(* IEC 61131-3 sources: plc-st-coding-agent/progress/evidence/f14_v14_remaining_20261113/jobs/codex_deepseek-v4pro (part 2) *)

(* ---- public-hard-01.raw_candidate_03.st ---- *)
(* CONTRACT_RULES [] *)

(* ENGINEERING_CONTRACT
   - ESTOP: ESTOP=FALSE forces every output OFF in this scan; manual and auto commands are inhibited.
   - Manual runs: only while OpeMode=FALSE and ESTOP=TRUE; each start button rising edge toggles its retained output latch.
   - Auto sequence: AUTOSTART rising edge while OpeMode=TRUE enters FILL_A; output valves follow the sequence below.
   - Valve A: ON in FILL_A; Level>=50 closes A and opens B (PUB012).
   - Valve B: ON in FILL_B; Level>=80 closes B (PUB012/PUB013).
   - ProcessMode=FALSE: at Level>=80 mixer starts; MixMotorComplete latches completion, then mixer off and Valve D ON, sequence done (PUB014).
   - ProcessMode=TRUE: at Level>=80 Valve C opens; Level>=100 closes C and starts mixer; completion opens D (PUB014).
   - Mix complete is latched until the next AUTOSTART; Valve D remains ON in DONE because no stop/reset is stated.
   - Thresholds are inclusive >=; Level is INT cm; PROCESSMODE is read live at the 80 cm transition.
*)

TYPE E_MaterialProportioningState :
(
    MP_IDLE,
    MP_FILL_A,
    MP_FILL_B,
    MP_MIX_SIMPLE,
    MP_FILL_C,
    MP_MIX_C,
    MP_DONE
) := MP_IDLE;
END_TYPE;

FUNCTION_BLOCK MaterialProportioningControl
VAR_INPUT
    estop : BOOL;
    opeMode : BOOL;
    valveAStart : BOOL;
    valveBStart : BOOL;
    valveCStart : BOOL;
    valveDStart : BOOL;
    mixMotorStart : BOOL;
    autoStart : BOOL;
    processMode : BOOL;
    levelSensor : INT;
    mixMotorComplete : BOOL;
END_VAR
VAR_OUTPUT
    valveARun : BOOL;
    valveBRun : BOOL;
    valveCRun : BOOL;
    valveDRun : BOOL;
    mixMotorRun : BOOL;
END_VAR
VAR
    tmp_trigValveA : R_TRIG;
    tmp_trigValveB : R_TRIG;
    tmp_trigValveC : R_TRIG;
    tmp_trigValveD : R_TRIG;
    tmp_trigMixMotor : R_TRIG;
    tmp_trigAutoStart : R_TRIG;

    manualValveARun : BOOL := FALSE;
    manualValveBRun : BOOL := FALSE;
    manualValveCRun : BOOL := FALSE;
    manualValveDRun : BOOL := FALSE;
    manualMixMotorRun : BOOL := FALSE;

    state : E_MaterialProportioningState := MP_IDLE;
    mixCompleteLatched : BOOL := FALSE;
END_VAR

tmp_trigValveA(CLK := valveAStart);
tmp_trigValveB(CLK := valveBStart);
tmp_trigValveC(CLK := valveCStart);
tmp_trigValveD(CLK := valveDStart);
tmp_trigMixMotor(CLK := mixMotorStart);
tmp_trigAutoStart(CLK := autoStart);

IF NOT estop THEN
    valveARun := FALSE;
    valveBRun := FALSE;
    valveCRun := FALSE;
    valveDRun := FALSE;
    mixMotorRun := FALSE;

ELSIF NOT opeMode THEN
    state := MP_IDLE;
    mixCompleteLatched := FALSE;

    IF tmp_trigValveA.Q THEN
        manualValveARun := NOT manualValveARun;
    END_IF;
    IF tmp_trigValveB.Q THEN
        manualValveBRun := NOT manualValveBRun;
    END_IF;
    IF tmp_trigValveC.Q THEN
        manualValveCRun := NOT manualValveCRun;
    END_IF;
    IF tmp_trigValveD.Q THEN
        manualValveDRun := NOT manualValveDRun;
    END_IF;
    IF tmp_trigMixMotor.Q THEN
        manualMixMotorRun := NOT manualMixMotorRun;
    END_IF;

    valveARun := manualValveARun;
    valveBRun := manualValveBRun;
    valveCRun := manualValveCRun;
    valveDRun := manualValveDRun;
    mixMotorRun := manualMixMotorRun;

ELSE
    IF tmp_trigAutoStart.Q THEN
        state := MP_FILL_A;
        mixCompleteLatched := FALSE;
    END_IF;

    CASE state OF
        MP_IDLE:
            valveARun := FALSE;
            valveBRun := FALSE;
            valveCRun := FALSE;
            valveDRun := FALSE;
            mixMotorRun := FALSE;

        MP_FILL_A:
            valveARun := TRUE;
            valveBRun := FALSE;
            valveCRun := FALSE;
            valveDRun := FALSE;
            mixMotorRun := FALSE;

            IF levelSensor >= 80 THEN
                valveARun := FALSE;
                valveBRun := FALSE;
                IF NOT processMode THEN
                    mixMotorRun := TRUE;
                    mixCompleteLatched := FALSE;
                    state := MP_MIX_SIMPLE;
                ELSIF levelSensor >= 100 THEN
                    valveCRun := FALSE;
                    mixMotorRun := TRUE;
                    mixCompleteLatched := FALSE;
                    state := MP_MIX_C;
                ELSE
                    valveCRun := TRUE;
                    state := MP_FILL_C;
                END_IF;
            ELSIF levelSensor >= 50 THEN
                valveARun := FALSE;
                valveBRun := TRUE;
                state := MP_FILL_B;
            END_IF;

        MP_FILL_B:
            valveARun := FALSE;
            valveBRun := TRUE;
            valveCRun := FALSE;
            valveDRun := FALSE;
            mixMotorRun := FALSE;

            IF levelSensor >= 80 THEN
                valveBRun := FALSE;
                IF NOT processMode THEN
                    mixMotorRun := TRUE;
                    mixCompleteLatched := FALSE;
                    state := MP_MIX_SIMPLE;
                ELSE
                    IF levelSensor >= 100 THEN
                        valveCRun := FALSE;
                        mixMotorRun := TRUE;
                        mixCompleteLatched := FALSE;
                        state := MP_MIX_C;
                    ELSE
                        valveCRun := TRUE;
                        state := MP_FILL_C;
                    END_IF;
                END_IF;
            END_IF;

        MP_FILL_C:
            valveARun := FALSE;
            valveBRun := FALSE;
            valveCRun := TRUE;
            valveDRun := FALSE;
            mixMotorRun := FALSE;

            IF levelSensor >= 100 THEN
                valveCRun := FALSE;
                mixMotorRun := TRUE;
                mixCompleteLatched := FALSE;
                state := MP_MIX_C;
            END_IF;

        MP_MIX_SIMPLE:
            valveARun := FALSE;
            valveBRun := FALSE;
            valveCRun := FALSE;
            valveDRun := FALSE;
            mixMotorRun := TRUE;

            IF mixMotorComplete THEN
                mixCompleteLatched := TRUE;
            END_IF;

            IF mixCompleteLatched THEN
                mixMotorRun := FALSE;
                valveDRun := TRUE;
                state := MP_DONE;
            END_IF;

        MP_MIX_C:
            valveARun := FALSE;
            valveBRun := FALSE;
            valveCRun := FALSE;
            valveDRun := FALSE;
            mixMotorRun := TRUE;

            IF mixMotorComplete THEN
                mixCompleteLatched := TRUE;
            END_IF;

            IF mixCompleteLatched THEN
                mixMotorRun := FALSE;
                valveDRun := TRUE;
                state := MP_DONE;
            END_IF;

        MP_DONE:
            valveARun := FALSE;
            valveBRun := FALSE;
            valveCRun := FALSE;
            valveDRun := TRUE;
            mixMotorRun := FALSE;
    END_CASE;
END_IF;
END_FUNCTION_BLOCK

(* ---- public-hard-02.candidate_01.st ---- *)
(*
ENGINEERING_CONTRACT
- conveyorLeft | activation: ST_MOVING and target<current | hold: while ST_MOVING | reset: target sensor arrival or non-moving state | same-scan: final settled state/target controls write | PUB001,PUB005.
- conveyorRight | activation: ST_MOVING and target>current | hold: while ST_MOVING | reset: target sensor arrival or non-moving state | same-scan: final settled state/target controls write | PUB001,PUB005.
- local_state | activation: ST_IDLE+start -> ST_MOVING; ST_MOVING+sensor -> ST_WAIT_COMPLETION/ST_DONE/next ST_MOVING; ST_WAIT_COMPLETION+completion -> ST_MOVING/ST_DONE | hold: retained every scan | reset/deactivation: above transitions | same-scan: inputs iterated to fixed point before outputs | units: seq index 1..processLength, stations 1..5 | PUB001-PUB005.
- local_step_index/current/target | update: start, sensor, completion | hold: otherwise | bounds: step 1..8, current/target 1..5 | PUB002,PUB005.
- Direction rule: one target per step yields exactly one direction output; equal/unknown target de-energizes both.
- Unspecified: no restart/reset after station5; completion signals treated as levels.
*)
(* CONTRACT_RULES [] *)

TYPE CONTROL_STATE :
(
    ST_IDLE,
    ST_MOVING,
    ST_WAIT_COMPLETION,
    ST_DONE
);
END_TYPE;

FUNCTION_BLOCK FlexibleProcessingControl
VAR_INPUT
    processLength : USINT;
    sensor1 : BOOL;
    sensor2 : BOOL;
    sensor3 : BOOL;
    sensor4 : BOOL;
    sensor5 : BOOL;
    station1Start : BOOL;
    station2Complete : BOOL;
    station3Complete : BOOL;
    station4Complete : BOOL;
    processSequence : ARRAY[1..8] OF USINT;
END_VAR
VAR_OUTPUT
    conveyorLeft : BOOL;
    conveyorRight : BOOL;
END_VAR
VAR
    local_state : CONTROL_STATE := ST_IDLE;
    local_step_index : USINT := 0;
    local_current_station : USINT := 1;
    local_target_station : USINT := 0;
    local_completion_active : BOOL := FALSE;
    local_target_sensor_active : BOOL := FALSE;
    local_fixpoint_scan : INT := 0;
    local_fixpoint_stable : BOOL := FALSE;
END_VAR

FOR local_fixpoint_scan := 1 TO 20 DO
    local_fixpoint_stable := TRUE;

    local_completion_active := FALSE;
    IF local_target_station = 2 THEN
        local_completion_active := station2Complete;
    ELSIF local_target_station = 3 THEN
        local_completion_active := station3Complete;
    ELSIF local_target_station = 4 THEN
        local_completion_active := station4Complete;
    END_IF;

    local_target_sensor_active := FALSE;
    IF local_target_station = 2 THEN
        local_target_sensor_active := sensor2;
    ELSIF local_target_station = 3 THEN
        local_target_sensor_active := sensor3;
    ELSIF local_target_station = 4 THEN
        local_target_sensor_active := sensor4;
    ELSIF local_target_station = 5 THEN
        local_target_sensor_active := sensor5;
    END_IF;

    CASE local_state OF
        ST_IDLE:
            IF sensor1 AND station1Start THEN
                local_step_index := 1;
                local_current_station := 1;
                local_target_station := processSequence[1];
                local_state := ST_MOVING;
                local_fixpoint_stable := FALSE;
            END_IF;

        ST_MOVING:
            IF local_target_sensor_active THEN
                local_current_station := local_target_station;

                IF local_target_station = 5 THEN
                    local_state := ST_DONE;
                ELSIF local_completion_active THEN
                    IF local_step_index < processLength THEN
                        local_step_index := local_step_index + 1;
                        local_target_station := processSequence[local_step_index];
                        local_state := ST_MOVING;
                    ELSE
                        local_state := ST_DONE;
                    END_IF;
                ELSE
                    local_state := ST_WAIT_COMPLETION;
                END_IF;

                local_fixpoint_stable := FALSE;
            END_IF;

        ST_WAIT_COMPLETION:
            IF local_completion_active THEN
                IF local_step_index < processLength THEN
                    local_step_index := local_step_index + 1;
                    local_target_station := processSequence[local_step_index];
                    local_state := ST_MOVING;
                ELSE
                    local_state := ST_DONE;
                END_IF;

                local_fixpoint_stable := FALSE;
            END_IF;

        ST_DONE:
            local_fixpoint_stable := TRUE;
    END_CASE;

    IF local_fixpoint_stable THEN
        EXIT;
    END_IF;
END_FOR;

IF local_state = ST_MOVING THEN
    IF local_target_station > local_current_station THEN
        conveyorLeft := FALSE;
        conveyorRight := TRUE;
    ELSIF local_target_station < local_current_station THEN
        conveyorLeft := TRUE;
        conveyorRight := FALSE;
    ELSE
        conveyorLeft := FALSE;
        conveyorRight := FALSE;
    END_IF;
ELSE
    conveyorLeft := FALSE;
    conveyorRight := FALSE;
END_IF;

END_FUNCTION_BLOCK

(* ---- public-hard-02.candidate_02.st ---- *)
(*
ENGINEERING_CONTRACT
- conveyorLeft | activation: ST_MOVING and target<current | hold: while ST_MOVING | reset: target sensor arrival or non-moving state | same-scan: final settled state/target controls write | PUB001,PUB005.
- conveyorRight | activation: ST_MOVING and target>current | hold: while ST_MOVING | reset: target sensor arrival or non-moving state | same-scan: final settled state/target controls write | PUB001,PUB005.
- local_state | activation: ST_IDLE+start -> ST_MOVING; ST_MOVING+sensor -> ST_WAIT_COMPLETION/ST_DONE/next ST_MOVING; ST_WAIT_COMPLETION+completion -> ST_MOVING/ST_DONE | hold: retained every scan | reset/deactivation: above transitions | same-scan: inputs iterated to fixed point before outputs | units: seq index 1..processLength, stations 1..5 | PUB001-PUB005.
- local_step_index/current/target | update: start, sensor, completion | hold: otherwise | bounds: step 1..8, current/target 1..5 | PUB002,PUB005.
- Direction rule: one target per step yields exactly one direction output; equal/unknown target de-energizes both.
- Unspecified: completion signals treated as levels; ST_DONE restarts on sensor1 AND station1Start.
*)
(* CONTRACT_RULES [] *)

TYPE CONTROL_STATE :
(
    ST_IDLE,
    ST_MOVING,
    ST_WAIT_COMPLETION,
    ST_DONE
);
END_TYPE;

FUNCTION_BLOCK FlexibleProcessingControl
VAR_INPUT
    processLength : USINT;
    sensor1 : BOOL;
    sensor2 : BOOL;
    sensor3 : BOOL;
    sensor4 : BOOL;
    sensor5 : BOOL;
    station1Start : BOOL;
    station2Complete : BOOL;
    station3Complete : BOOL;
    station4Complete : BOOL;
    processSequence : ARRAY[1..8] OF USINT;
END_VAR
VAR_OUTPUT
    conveyorLeft : BOOL;
    conveyorRight : BOOL;
END_VAR
VAR
    local_state : CONTROL_STATE := ST_IDLE;
    local_step_index : USINT := 0;
    local_current_station : USINT := 1;
    local_target_station : USINT := 0;
    local_completion_active : BOOL := FALSE;
    local_target_sensor_active : BOOL := FALSE;
    local_fixpoint_scan : INT := 0;
    local_fixpoint_stable : BOOL := FALSE;
END_VAR

FOR local_fixpoint_scan := 1 TO 20 DO
    local_fixpoint_stable := TRUE;

    local_completion_active := FALSE;
    IF local_target_station = 2 THEN
        local_completion_active := station2Complete;
    ELSIF local_target_station = 3 THEN
        local_completion_active := station3Complete;
    ELSIF local_target_station = 4 THEN
        local_completion_active := station4Complete;
    END_IF;

    local_target_sensor_active := FALSE;
    IF local_target_station = 2 THEN
        local_target_sensor_active := sensor2;
    ELSIF local_target_station = 3 THEN
        local_target_sensor_active := sensor3;
    ELSIF local_target_station = 4 THEN
        local_target_sensor_active := sensor4;
    ELSIF local_target_station = 5 THEN
        local_target_sensor_active := sensor5;
    END_IF;

    CASE local_state OF
        ST_IDLE:
            IF sensor1 AND station1Start THEN
                local_step_index := 1;
                local_current_station := 1;
                local_target_station := processSequence[1];
                local_state := ST_MOVING;
                local_fixpoint_stable := FALSE;
            END_IF;

        ST_MOVING:
            IF local_target_sensor_active THEN
                local_current_station := local_target_station;

                IF local_target_station = 5 THEN
                    local_state := ST_DONE;
                ELSIF local_completion_active THEN
                    IF local_step_index < processLength THEN
                        local_step_index := local_step_index + 1;
                        local_target_station := processSequence[local_step_index];
                        local_state := ST_MOVING;
                    ELSE
                        local_state := ST_DONE;
                    END_IF;
                ELSE
                    local_state := ST_WAIT_COMPLETION;
                END_IF;

                local_fixpoint_stable := FALSE;
            END_IF;

        ST_WAIT_COMPLETION:
            IF local_completion_active THEN
                IF local_step_index < processLength THEN
                    local_step_index := local_step_index + 1;
                    local_target_station := processSequence[local_step_index];
                    local_state := ST_MOVING;
                ELSE
                    local_state := ST_DONE;
                END_IF;

                local_fixpoint_stable := FALSE;
            END_IF;

        ST_DONE:
            IF sensor1 AND station1Start THEN
                local_step_index := 1;
                local_current_station := 1;
                local_target_station := processSequence[1];
                local_state := ST_MOVING;
                local_fixpoint_stable := FALSE;
            END_IF;
    END_CASE;

    IF local_fixpoint_stable THEN
        EXIT;
    END_IF;
END_FOR;

IF local_state = ST_MOVING THEN
    IF local_target_station > local_current_station THEN
        conveyorLeft := FALSE;
        conveyorRight := TRUE;
    ELSIF local_target_station < local_current_station THEN
        conveyorLeft := TRUE;
        conveyorRight := FALSE;
    ELSE
        conveyorLeft := FALSE;
        conveyorRight := FALSE;
    END_IF;
ELSE
    conveyorLeft := FALSE;
    conveyorRight := FALSE;
END_IF;

END_FUNCTION_BLOCK

(* ---- public-hard-02.candidate_03.st ---- *)
(*
ENGINEERING_CONTRACT
- conveyorLeft | activation: ST_MOVING and target<current | hold: while ST_MOVING | reset: target sensor arrival or non-moving state | same-scan: final settled state/target controls write | PUB001,PUB005.
- conveyorRight | activation: ST_MOVING and target>current | hold: while ST_MOVING | reset: target sensor arrival or non-moving state | same-scan: final settled state/target controls write | PUB001,PUB005.
- local_state | activation: ST_IDLE+start -> ST_MOVING; ST_MOVING+sensor -> ST_WAIT_COMPLETION/ST_DONE/next ST_MOVING; ST_WAIT_COMPLETION+completion -> ST_MOVING/ST_DONE | hold: retained every scan | reset/deactivation: above transitions | same-scan: one transition per scan based on current public inputs | units: seq index 1..processLength, stations 1..5 | PUB001-PUB005.
- local_step_index/current/target | update: start, sensor, completion | hold: otherwise | bounds: step 1..8, current/target 1..5 | PUB002,PUB005.
- Direction rule: one target per step yields exactly one direction output; equal/unknown target de-energizes both.
- Unspecified: completion signals treated as levels; ST_DONE restarts on sensor1 AND station1Start.
*)
(* CONTRACT_RULES [] *)

TYPE CONTROL_STATE :
(
    ST_IDLE,
    ST_MOVING,
    ST_WAIT_COMPLETION,
    ST_DONE
);
END_TYPE;

FUNCTION_BLOCK FlexibleProcessingControl
VAR_INPUT
    processLength : USINT;
    sensor1 : BOOL;
    sensor2 : BOOL;
    sensor3 : BOOL;
    sensor4 : BOOL;
    sensor5 : BOOL;
    station1Start : BOOL;
    station2Complete : BOOL;
    station3Complete : BOOL;
    station4Complete : BOOL;
    processSequence : ARRAY[1..8] OF USINT;
END_VAR
VAR_OUTPUT
    conveyorLeft : BOOL;
    conveyorRight : BOOL;
END_VAR
VAR
    local_state : CONTROL_STATE := ST_IDLE;
    local_step_index : USINT := 0;
    local_current_station : USINT := 1;
    local_target_station : USINT := 0;
    local_completion_active : BOOL := FALSE;
    local_target_sensor_active : BOOL := FALSE;
END_VAR

    local_completion_active := FALSE;
    IF local_target_station = 2 THEN
        local_completion_active := station2Complete;
    ELSIF local_target_station = 3 THEN
        local_completion_active := station3Complete;
    ELSIF local_target_station = 4 THEN
        local_completion_active := station4Complete;
    END_IF;

    local_target_sensor_active := FALSE;
    IF local_target_station = 2 THEN
        local_target_sensor_active := sensor2;
    ELSIF local_target_station = 3 THEN
        local_target_sensor_active := sensor3;
    ELSIF local_target_station = 4 THEN
        local_target_sensor_active := sensor4;
    ELSIF local_target_station = 5 THEN
        local_target_sensor_active := sensor5;
    END_IF;

    CASE local_state OF
        ST_IDLE:
            IF sensor1 AND station1Start THEN
                local_step_index := 1;
                local_current_station := 1;
                local_target_station := processSequence[1];
                local_state := ST_MOVING;
            END_IF;

        ST_MOVING:
            IF local_target_sensor_active THEN
                local_current_station := local_target_station;

                IF local_target_station = 5 THEN
                    local_state := ST_DONE;
                ELSIF local_completion_active THEN
                    IF local_step_index < processLength THEN
                        local_step_index := local_step_index + 1;
                        local_target_station := processSequence[local_step_index];
                        local_state := ST_MOVING;
                    ELSE
                        local_state := ST_DONE;
                    END_IF;
                ELSE
                    local_state := ST_WAIT_COMPLETION;
                END_IF;
            END_IF;

        ST_WAIT_COMPLETION:
            IF local_completion_active THEN
                IF local_step_index < processLength THEN
                    local_step_index := local_step_index + 1;
                    local_target_station := processSequence[local_step_index];
                    local_state := ST_MOVING;
                ELSE
                    local_state := ST_DONE;
                END_IF;
            END_IF;

        ST_DONE:
            IF sensor1 AND station1Start THEN
                local_step_index := 1;
                local_current_station := 1;
                local_target_station := processSequence[1];
                local_state := ST_MOVING;
            END_IF;
    END_CASE;

IF local_state = ST_MOVING THEN
    IF local_target_station > local_current_station THEN
        conveyorLeft := FALSE;
        conveyorRight := TRUE;
    ELSIF local_target_station < local_current_station THEN
        conveyorLeft := TRUE;
        conveyorRight := FALSE;
    ELSE
        conveyorLeft := FALSE;
        conveyorRight := FALSE;
    END_IF;
ELSE
    conveyorLeft := FALSE;
    conveyorRight := FALSE;
END_IF;

END_FUNCTION_BLOCK

(* ---- public-hard-02.patch_base_02.st ---- *)
(*
ENGINEERING_CONTRACT
- conveyorLeft | activation: ST_MOVING and target<current | hold: while ST_MOVING | reset: target sensor arrival or non-moving state | same-scan: final settled state/target controls write | PUB001,PUB005.
- conveyorRight | activation: ST_MOVING and target>current | hold: while ST_MOVING | reset: target sensor arrival or non-moving state | same-scan: final settled state/target controls write | PUB001,PUB005.
- local_state | activation: ST_IDLE+start -> ST_MOVING; ST_MOVING+sensor -> ST_WAIT_COMPLETION/ST_DONE/next ST_MOVING; ST_WAIT_COMPLETION+completion -> ST_MOVING/ST_DONE | hold: retained every scan | reset/deactivation: above transitions | same-scan: inputs iterated to fixed point before outputs | units: seq index 1..processLength, stations 1..5 | PUB001-PUB005.
- local_step_index/current/target | update: start, sensor, completion | hold: otherwise | bounds: step 1..8, current/target 1..5 | PUB002,PUB005.
- Direction rule: one target per step yields exactly one direction output; equal/unknown target de-energizes both.
- Unspecified: no restart/reset after station5; completion signals treated as levels.
*)
(* CONTRACT_RULES [] *)

TYPE CONTROL_STATE :
(
    ST_IDLE,
    ST_MOVING,
    ST_WAIT_COMPLETION,
    ST_DONE
);
END_TYPE;

FUNCTION_BLOCK FlexibleProcessingControl
VAR_INPUT
    processLength : USINT;
    sensor1 : BOOL;
    sensor2 : BOOL;
    sensor3 : BOOL;
    sensor4 : BOOL;
    sensor5 : BOOL;
    station1Start : BOOL;
    station2Complete : BOOL;
    station3Complete : BOOL;
    station4Complete : BOOL;
    processSequence : ARRAY[1..8] OF USINT;
END_VAR
VAR_OUTPUT
    conveyorLeft : BOOL;
    conveyorRight : BOOL;
END_VAR
VAR
    local_state : CONTROL_STATE := ST_IDLE;
    local_step_index : USINT := 0;
    local_current_station : USINT := 1;
    local_target_station : USINT := 0;
    local_completion_active : BOOL := FALSE;
    local_target_sensor_active : BOOL := FALSE;
    local_fixpoint_scan : INT := 0;
    local_fixpoint_stable : BOOL := FALSE;
END_VAR

FOR local_fixpoint_scan := 1 TO 20 DO
    local_fixpoint_stable := TRUE;

    local_completion_active := FALSE;
    IF local_target_station = 2 THEN
        local_completion_active := station2Complete;
    ELSIF local_target_station = 3 THEN
        local_completion_active := station3Complete;
    ELSIF local_target_station = 4 THEN
        local_completion_active := station4Complete;
    END_IF;

    local_target_sensor_active := FALSE;
    IF local_target_station = 2 THEN
        local_target_sensor_active := sensor2;
    ELSIF local_target_station = 3 THEN
        local_target_sensor_active := sensor3;
    ELSIF local_target_station = 4 THEN
        local_target_sensor_active := sensor4;
    ELSIF local_target_station = 5 THEN
        local_target_sensor_active := sensor5;
    END_IF;

    CASE local_state OF
        ST_IDLE:
            IF sensor1 AND station1Start THEN
                local_step_index := 1;
                local_current_station := 1;
                local_target_station := processSequence[1];
                local_state := ST_MOVING;
                local_fixpoint_stable := FALSE;
            END_IF;

        ST_MOVING:
            IF local_target_sensor_active THEN
                local_current_station := local_target_station;

                IF local_target_station = 5 THEN
                    local_state := ST_DONE;
                ELSIF local_completion_active THEN
                    IF local_step_index < processLength THEN
                        local_step_index := local_step_index + 1;
                        local_target_station := processSequence[local_step_index];
                        local_state := ST_MOVING;
                    ELSE
                        local_state := ST_DONE;
                    END_IF;
                ELSE
                    local_state := ST_WAIT_COMPLETION;
                END_IF;

                local_fixpoint_stable := FALSE;
            END_IF;

        ST_WAIT_COMPLETION:
            IF local_completion_active THEN
                IF local_step_index < processLength THEN
                    local_step_index := local_step_index + 1;
                    local_target_station := processSequence[local_step_index];
                    local_state := ST_MOVING;
                ELSE
                    local_state := ST_DONE;
                END_IF;

                local_fixpoint_stable := FALSE;
            END_IF;

        ST_DONE:
            local_fixpoint_stable := TRUE;
    END_CASE;

    IF local_fixpoint_stable THEN
        EXIT;
    END_IF;
END_FOR;

IF local_state = ST_MOVING THEN
    IF local_target_station > local_current_station THEN
        conveyorLeft := FALSE;
        conveyorRight := TRUE;
    ELSIF local_target_station < local_current_station THEN
        conveyorLeft := TRUE;
        conveyorRight := FALSE;
    ELSE
        conveyorLeft := FALSE;
        conveyorRight := FALSE;
    END_IF;
ELSE
    conveyorLeft := FALSE;
    conveyorRight := FALSE;
END_IF;

END_FUNCTION_BLOCK

(* ---- public-hard-02.patch_base_03.st ---- *)
(*
ENGINEERING_CONTRACT
- conveyorLeft | activation: ST_MOVING and target<current | hold: while ST_MOVING | reset: target sensor arrival or non-moving state | same-scan: final settled state/target controls write | PUB001,PUB005.
- conveyorRight | activation: ST_MOVING and target>current | hold: while ST_MOVING | reset: target sensor arrival or non-moving state | same-scan: final settled state/target controls write | PUB001,PUB005.
- local_state | activation: ST_IDLE+start -> ST_MOVING; ST_MOVING+sensor -> ST_WAIT_COMPLETION/ST_DONE/next ST_MOVING; ST_WAIT_COMPLETION+completion -> ST_MOVING/ST_DONE | hold: retained every scan | reset/deactivation: above transitions | same-scan: inputs iterated to fixed point before outputs | units: seq index 1..processLength, stations 1..5 | PUB001-PUB005.
- local_step_index/current/target | update: start, sensor, completion | hold: otherwise | bounds: step 1..8, current/target 1..5 | PUB002,PUB005.
- Direction rule: one target per step yields exactly one direction output; equal/unknown target de-energizes both.
- Unspecified: completion signals treated as levels; ST_DONE restarts on sensor1 AND station1Start.
*)
(* CONTRACT_RULES [] *)

TYPE CONTROL_STATE :
(
    ST_IDLE,
    ST_MOVING,
    ST_WAIT_COMPLETION,
    ST_DONE
);
END_TYPE;

FUNCTION_BLOCK FlexibleProcessingControl
VAR_INPUT
    processLength : USINT;
    sensor1 : BOOL;
    sensor2 : BOOL;
    sensor3 : BOOL;
    sensor4 : BOOL;
    sensor5 : BOOL;
    station1Start : BOOL;
    station2Complete : BOOL;
    station3Complete : BOOL;
    station4Complete : BOOL;
    processSequence : ARRAY[1..8] OF USINT;
END_VAR
VAR_OUTPUT
    conveyorLeft : BOOL;
    conveyorRight : BOOL;
END_VAR
VAR
    local_state : CONTROL_STATE := ST_IDLE;
    local_step_index : USINT := 0;
    local_current_station : USINT := 1;
    local_target_station : USINT := 0;
    local_completion_active : BOOL := FALSE;
    local_target_sensor_active : BOOL := FALSE;
    local_fixpoint_scan : INT := 0;
    local_fixpoint_stable : BOOL := FALSE;
END_VAR

FOR local_fixpoint_scan := 1 TO 20 DO
    local_fixpoint_stable := TRUE;

    local_completion_active := FALSE;
    IF local_target_station = 2 THEN
        local_completion_active := station2Complete;
    ELSIF local_target_station = 3 THEN
        local_completion_active := station3Complete;
    ELSIF local_target_station = 4 THEN
        local_completion_active := station4Complete;
    END_IF;

    local_target_sensor_active := FALSE;
    IF local_target_station = 2 THEN
        local_target_sensor_active := sensor2;
    ELSIF local_target_station = 3 THEN
        local_target_sensor_active := sensor3;
    ELSIF local_target_station = 4 THEN
        local_target_sensor_active := sensor4;
    ELSIF local_target_station = 5 THEN
        local_target_sensor_active := sensor5;
    END_IF;

    CASE local_state OF
        ST_IDLE:
            IF sensor1 AND station1Start THEN
                local_step_index := 1;
                local_current_station := 1;
                local_target_station := processSequence[1];
                local_state := ST_MOVING;
                local_fixpoint_stable := FALSE;
            END_IF;

        ST_MOVING:
            IF local_target_sensor_active THEN
                local_current_station := local_target_station;

                IF local_target_station = 5 THEN
                    local_state := ST_DONE;
                ELSIF local_completion_active THEN
                    IF local_step_index < processLength THEN
                        local_step_index := local_step_index + 1;
                        local_target_station := processSequence[local_step_index];
                        local_state := ST_MOVING;
                    ELSE
                        local_state := ST_DONE;
                    END_IF;
                ELSE
                    local_state := ST_WAIT_COMPLETION;
                END_IF;

                local_fixpoint_stable := FALSE;
            END_IF;

        ST_WAIT_COMPLETION:
            IF local_completion_active THEN
                IF local_step_index < processLength THEN
                    local_step_index := local_step_index + 1;
                    local_target_station := processSequence[local_step_index];
                    local_state := ST_MOVING;
                ELSE
                    local_state := ST_DONE;
                END_IF;

                local_fixpoint_stable := FALSE;
            END_IF;

        ST_DONE:
            IF sensor1 AND station1Start THEN
                local_step_index := 1;
                local_current_station := 1;
                local_target_station := processSequence[1];
                local_state := ST_MOVING;
                local_fixpoint_stable := FALSE;
            END_IF;
    END_CASE;

    IF local_fixpoint_stable THEN
        EXIT;
    END_IF;
END_FOR;

IF local_state = ST_MOVING THEN
    IF local_target_station > local_current_station THEN
        conveyorLeft := FALSE;
        conveyorRight := TRUE;
    ELSIF local_target_station < local_current_station THEN
        conveyorLeft := TRUE;
        conveyorRight := FALSE;
    ELSE
        conveyorLeft := FALSE;
        conveyorRight := FALSE;
    END_IF;
ELSE
    conveyorLeft := FALSE;
    conveyorRight := FALSE;
END_IF;

END_FUNCTION_BLOCK

(* ---- public-hard-02.raw_candidate_01.st ---- *)
(*
ENGINEERING_CONTRACT
- conveyorLeft | activation: ST_MOVING and target<current | hold: while ST_MOVING | reset: target sensor arrival or non-moving state | same-scan: final settled state/target controls write | PUB001,PUB005.
- conveyorRight | activation: ST_MOVING and target>current | hold: while ST_MOVING | reset: target sensor arrival or non-moving state | same-scan: final settled state/target controls write | PUB001,PUB005.
- local_state | activation: ST_IDLE+start -> ST_MOVING; ST_MOVING+sensor -> ST_WAIT_COMPLETION/ST_DONE/next ST_MOVING; ST_WAIT_COMPLETION+completion -> ST_MOVING/ST_DONE | hold: retained every scan | reset/deactivation: above transitions | same-scan: inputs iterated to fixed point before outputs | units: seq index 1..processLength, stations 1..5 | PUB001-PUB005.
- local_step_index/current/target | update: start, sensor, completion | hold: otherwise | bounds: step 1..8, current/target 1..5 | PUB002,PUB005.
- Direction rule: one target per step yields exactly one direction output; equal/unknown target de-energizes both.
- Unspecified: no restart/reset after station5; completion signals treated as levels.
*)
(* CONTRACT_RULES [] *)

TYPE CONTROL_STATE :
(
    ST_IDLE,
    ST_MOVING,
    ST_WAIT_COMPLETION,
    ST_DONE
);
END_TYPE

FUNCTION_BLOCK FlexibleProcessingControl
VAR_INPUT
    processLength : USINT;
    sensor1 : BOOL;
    sensor2 : BOOL;
    sensor3 : BOOL;
    sensor4 : BOOL;
    sensor5 : BOOL;
    station1Start : BOOL;
    station2Complete : BOOL;
    station3Complete : BOOL;
    station4Complete : BOOL;
    processSequence : ARRAY[1..8] OF USINT;
END_VAR
VAR_OUTPUT
    conveyorLeft : BOOL;
    conveyorRight : BOOL;
END_VAR
VAR
    local_state : CONTROL_STATE := ST_IDLE;
    local_step_index : USINT := 0;
    local_current_station : USINT := 1;
    local_target_station : USINT := 0;
    local_completion_active : BOOL := FALSE;
    local_target_sensor_active : BOOL := FALSE;
    local_fixpoint_scan : INT := 0;
    local_fixpoint_stable : BOOL := FALSE;
END_VAR

FOR local_fixpoint_scan := 1 TO 20 DO
    local_fixpoint_stable := TRUE;

    local_completion_active := FALSE;
    IF local_target_station = 2 THEN
        local_completion_active := station2Complete;
    ELSIF local_target_station = 3 THEN
        local_completion_active := station3Complete;
    ELSIF local_target_station = 4 THEN
        local_completion_active := station4Complete;
    END_IF;

    local_target_sensor_active := FALSE;
    IF local_target_station = 2 THEN
        local_target_sensor_active := sensor2;
    ELSIF local_target_station = 3 THEN
        local_target_sensor_active := sensor3;
    ELSIF local_target_station = 4 THEN
        local_target_sensor_active := sensor4;
    ELSIF local_target_station = 5 THEN
        local_target_sensor_active := sensor5;
    END_IF;

    CASE local_state OF
        ST_IDLE:
            IF sensor1 AND station1Start THEN
                local_step_index := 1;
                local_current_station := 1;
                local_target_station := processSequence[1];
                local_state := ST_MOVING;
                local_fixpoint_stable := FALSE;
            END_IF;

        ST_MOVING:
            IF local_target_sensor_active THEN
                local_current_station := local_target_station;

                IF local_target_station = 5 THEN
                    local_state := ST_DONE;
                ELSIF local_completion_active THEN
                    IF local_step_index < processLength THEN
                        local_step_index := local_step_index + 1;
                        local_target_station := processSequence[local_step_index];
                        local_state := ST_MOVING;
                    ELSE
                        local_state := ST_DONE;
                    END_IF;
                ELSE
                    local_state := ST_WAIT_COMPLETION;
                END_IF;

                local_fixpoint_stable := FALSE;
            END_IF;

        ST_WAIT_COMPLETION:
            IF local_completion_active THEN
                IF local_step_index < processLength THEN
                    local_step_index := local_step_index + 1;
                    local_target_station := processSequence[local_step_index];
                    local_state := ST_MOVING;
                ELSE
                    local_state := ST_DONE;
                END_IF;

                local_fixpoint_stable := FALSE;
            END_IF;

        ST_DONE:
            local_fixpoint_stable := TRUE;
    END_CASE;

    IF local_fixpoint_stable THEN
        EXIT;
    END_IF;
END_FOR;

IF local_state = ST_MOVING THEN
    IF local_target_station > local_current_station THEN
        conveyorLeft := FALSE;
        conveyorRight := TRUE;
    ELSIF local_target_station < local_current_station THEN
        conveyorLeft := TRUE;
        conveyorRight := FALSE;
    ELSE
        conveyorLeft := FALSE;
        conveyorRight := FALSE;
    END_IF;
ELSE
    conveyorLeft := FALSE;
    conveyorRight := FALSE;
END_IF;

END_FUNCTION_BLOCK

(* ---- public-hard-02.raw_candidate_02.st ---- *)
(*
ENGINEERING_CONTRACT
- conveyorLeft | activation: ST_MOVING and target<current | hold: while ST_MOVING | reset: target sensor arrival or non-moving state | same-scan: final settled state/target controls write | PUB001,PUB005.
- conveyorRight | activation: ST_MOVING and target>current | hold: while ST_MOVING | reset: target sensor arrival or non-moving state | same-scan: final settled state/target controls write | PUB001,PUB005.
- local_state | activation: ST_IDLE+start -> ST_MOVING; ST_MOVING+sensor -> ST_WAIT_COMPLETION/ST_DONE/next ST_MOVING; ST_WAIT_COMPLETION+completion -> ST_MOVING/ST_DONE | hold: retained every scan | reset/deactivation: above transitions | same-scan: inputs iterated to fixed point before outputs | units: seq index 1..processLength, stations 1..5 | PUB001-PUB005.
- local_step_index/current/target | update: start, sensor, completion | hold: otherwise | bounds: step 1..8, current/target 1..5 | PUB002,PUB005.
- Direction rule: one target per step yields exactly one direction output; equal/unknown target de-energizes both.
- Unspecified: completion signals treated as levels; ST_DONE restarts on sensor1 AND station1Start.
*)
(* CONTRACT_RULES [] *)

TYPE CONTROL_STATE :
(
    ST_IDLE,
    ST_MOVING,
    ST_WAIT_COMPLETION,
    ST_DONE
);
END_TYPE;

FUNCTION_BLOCK FlexibleProcessingControl
VAR_INPUT
    processLength : USINT;
    sensor1 : BOOL;
    sensor2 : BOOL;
    sensor3 : BOOL;
    sensor4 : BOOL;
    sensor5 : BOOL;
    station1Start : BOOL;
    station2Complete : BOOL;
    station3Complete : BOOL;
    station4Complete : BOOL;
    processSequence : ARRAY[1..8] OF USINT;
END_VAR
VAR_OUTPUT
    conveyorLeft : BOOL;
    conveyorRight : BOOL;
END_VAR
VAR
    local_state : CONTROL_STATE := ST_IDLE;
    local_step_index : USINT := 0;
    local_current_station : USINT := 1;
    local_target_station : USINT := 0;
    local_completion_active : BOOL := FALSE;
    local_target_sensor_active : BOOL := FALSE;
    local_fixpoint_scan : INT := 0;
    local_fixpoint_stable : BOOL := FALSE;
END_VAR

FOR local_fixpoint_scan := 1 TO 20 DO
    local_fixpoint_stable := TRUE;

    local_completion_active := FALSE;
    IF local_target_station = 2 THEN
        local_completion_active := station2Complete;
    ELSIF local_target_station = 3 THEN
        local_completion_active := station3Complete;
    ELSIF local_target_station = 4 THEN
        local_completion_active := station4Complete;
    END_IF;

    local_target_sensor_active := FALSE;
    IF local_target_station = 2 THEN
        local_target_sensor_active := sensor2;
    ELSIF local_target_station = 3 THEN
        local_target_sensor_active := sensor3;
    ELSIF local_target_station = 4 THEN
        local_target_sensor_active := sensor4;
    ELSIF local_target_station = 5 THEN
        local_target_sensor_active := sensor5;
    END_IF;

    CASE local_state OF
        ST_IDLE:
            IF sensor1 AND station1Start THEN
                local_step_index := 1;
                local_current_station := 1;
                local_target_station := processSequence[1];
                local_state := ST_MOVING;
                local_fixpoint_stable := FALSE;
            END_IF;

        ST_MOVING:
            IF local_target_sensor_active THEN
                local_current_station := local_target_station;

                IF local_target_station = 5 THEN
                    local_state := ST_DONE;
                ELSIF local_completion_active THEN
                    IF local_step_index < processLength THEN
                        local_step_index := local_step_index + 1;
                        local_target_station := processSequence[local_step_index];
                        local_state := ST_MOVING;
                    ELSE
                        local_state := ST_DONE;
                    END_IF;
                ELSE
                    local_state := ST_WAIT_COMPLETION;
                END_IF;

                local_fixpoint_stable := FALSE;
            END_IF;

        ST_WAIT_COMPLETION:
            IF local_completion_active THEN
                IF local_step_index < processLength THEN
                    local_step_index := local_step_index + 1;
                    local_target_station := processSequence[local_step_index];
                    local_state := ST_MOVING;
                ELSE
                    local_state := ST_DONE;
                END_IF;

                local_fixpoint_stable := FALSE;
            END_IF;

        ST_DONE:
            IF sensor1 AND station1Start THEN
                local_step_index := 1;
                local_current_station := 1;
                local_target_station := processSequence[1];
                local_state := ST_MOVING;
                local_fixpoint_stable := FALSE;
            END_IF;
    END_CASE;

    IF local_fixpoint_stable THEN
        EXIT;
    END_IF;
END_FOR;

IF local_state = ST_MOVING THEN
    IF local_target_station > local_current_station THEN
        conveyorLeft := FALSE;
        conveyorRight := TRUE;
    ELSIF local_target_station < local_current_station THEN
        conveyorLeft := TRUE;
        conveyorRight := FALSE;
    ELSE
        conveyorLeft := FALSE;
        conveyorRight := FALSE;
    END_IF;
ELSE
    conveyorLeft := FALSE;
    conveyorRight := FALSE;
END_IF;

END_FUNCTION_BLOCK

(* ---- public-hard-02.raw_candidate_03.st ---- *)
(*
ENGINEERING_CONTRACT
- conveyorLeft | activation: ST_MOVING and target<current | hold: while ST_MOVING | reset: target sensor arrival or non-moving state | same-scan: final settled state/target controls write | PUB001,PUB005.
- conveyorRight | activation: ST_MOVING and target>current | hold: while ST_MOVING | reset: target sensor arrival or non-moving state | same-scan: final settled state/target controls write | PUB001,PUB005.
- local_state | activation: ST_IDLE+start -> ST_MOVING; ST_MOVING+sensor -> ST_WAIT_COMPLETION/ST_DONE/next ST_MOVING; ST_WAIT_COMPLETION+completion -> ST_MOVING/ST_DONE | hold: retained every scan | reset/deactivation: above transitions | same-scan: one transition per scan based on current public inputs | units: seq index 1..processLength, stations 1..5 | PUB001-PUB005.
- local_step_index/current/target | update: start, sensor, completion | hold: otherwise | bounds: step 1..8, current/target 1..5 | PUB002,PUB005.
- Direction rule: one target per step yields exactly one direction output; equal/unknown target de-energizes both.
- Unspecified: completion signals treated as levels; ST_DONE restarts on sensor1 AND station1Start.
*)
(* CONTRACT_RULES [] *)

TYPE CONTROL_STATE :
(
    ST_IDLE,
    ST_MOVING,
    ST_WAIT_COMPLETION,
    ST_DONE
);
END_TYPE;

FUNCTION_BLOCK FlexibleProcessingControl
VAR_INPUT
    processLength : USINT;
    sensor1 : BOOL;
    sensor2 : BOOL;
    sensor3 : BOOL;
    sensor4 : BOOL;
    sensor5 : BOOL;
    station1Start : BOOL;
    station2Complete : BOOL;
    station3Complete : BOOL;
    station4Complete : BOOL;
    processSequence : ARRAY[1..8] OF USINT;
END_VAR
VAR_OUTPUT
    conveyorLeft : BOOL;
    conveyorRight : BOOL;
END_VAR
VAR
    local_state : CONTROL_STATE := ST_IDLE;
    local_step_index : USINT := 0;
    local_current_station : USINT := 1;
    local_target_station : USINT := 0;
    local_completion_active : BOOL := FALSE;
    local_target_sensor_active : BOOL := FALSE;
END_VAR

    local_completion_active := FALSE;
    IF local_target_station = 2 THEN
        local_completion_active := station2Complete;
    ELSIF local_target_station = 3 THEN
        local_completion_active := station3Complete;
    ELSIF local_target_station = 4 THEN
        local_completion_active := station4Complete;
    END_IF;

    local_target_sensor_active := FALSE;
    IF local_target_station = 2 THEN
        local_target_sensor_active := sensor2;
    ELSIF local_target_station = 3 THEN
        local_target_sensor_active := sensor3;
    ELSIF local_target_station = 4 THEN
        local_target_sensor_active := sensor4;
    ELSIF local_target_station = 5 THEN
        local_target_sensor_active := sensor5;
    END_IF;

    CASE local_state OF
        ST_IDLE:
            IF sensor1 AND station1Start THEN
                local_step_index := 1;
                local_current_station := 1;
                local_target_station := processSequence[1];
                local_state := ST_MOVING;
            END_IF;

        ST_MOVING:
            IF local_target_sensor_active THEN
                local_current_station := local_target_station;

                IF local_target_station = 5 THEN
                    local_state := ST_DONE;
                ELSIF local_completion_active THEN
                    IF local_step_index < processLength THEN
                        local_step_index := local_step_index + 1;
                        local_target_station := processSequence[local_step_index];
                        local_state := ST_MOVING;
                    ELSE
                        local_state := ST_DONE;
                    END_IF;
                ELSE
                    local_state := ST_WAIT_COMPLETION;
                END_IF;
            END_IF;

        ST_WAIT_COMPLETION:
            IF local_completion_active THEN
                IF local_step_index < processLength THEN
                    local_step_index := local_step_index + 1;
                    local_target_station := processSequence[local_step_index];
                    local_state := ST_MOVING;
                ELSE
                    local_state := ST_DONE;
                END_IF;
            END_IF;

        ST_DONE:
            IF sensor1 AND station1Start THEN
                local_step_index := 1;
                local_current_station := 1;
                local_target_station := processSequence[1];
                local_state := ST_MOVING;
            END_IF;
    END_CASE;

IF local_state = ST_MOVING THEN
    IF local_target_station > local_current_station THEN
        conveyorLeft := FALSE;
        conveyorRight := TRUE;
    ELSIF local_target_station < local_current_station THEN
        conveyorLeft := TRUE;
        conveyorRight := FALSE;
    ELSE
        conveyorLeft := FALSE;
        conveyorRight := FALSE;
    END_IF;
ELSE
    conveyorLeft := FALSE;
    conveyorRight := FALSE;
END_IF;

END_FUNCTION_BLOCK

(* ---- public-hard-03.candidate_01.st ---- *)
TYPE ST_Recipe :
STRUCT
    recipeID : INT;
    ingredientType : INT;
    ingredientRatio : REAL;
    productionTemperature : REAL;
END_STRUCT
END_TYPE;

FUNCTION_BLOCK FB_RecipeManagementSystem
VAR_INPUT
    addRecipe : BOOL;
    deleteRecipe : BOOL;
    modifyRecipe : BOOL;
    queryRecipe : BOOL;
    recipeIn : ST_Recipe;
END_VAR
VAR_OUTPUT
    recipeAdded : BOOL;
    recipeDeleted : BOOL;
    recipeModified : BOOL;
    recipeQueryResult : ST_Recipe;
    error : BOOL;
    status : WORD;
END_VAR
VAR_IN_OUT
    recipe : ARRAY[1..10] OF ST_Recipe;
END_VAR
VAR
    tmp_i : INT;
    tmp_foundIndex : INT;
    tmp_emptyIndex : INT;
    tmp_duplicateFound : BOOL;
    tmp_commandCount : INT;
    tmp_blankRecipe : ST_Recipe;
END_VAR

(* ENGINEERING_CONTRACT
   recipeAdded/Deleted/Modified: pulse TRUE only in the scan of a successful sole command; no retention; cleared each scan.
   recipeQueryResult: assigned from the matched recipe on a successful sole query; cleared to blank on all other scans; no retention.
   error/status: combinational per scan; PUB002-PUB006 error codes 16#8001..16#8005 on sole-command failures; 16#0000 on success/no operation.
   database recipe: retained through IN_OUT; altered only by successful add/delete/modify per PUB003-PUB005; slot recipeID=0 means empty.
   same-scan priority: simultaneous command requests are reported as unsupported with 16#8000; PUB011 leaves this case unspecified.
   units/boundaries: identifiers INT, ratios/temperatures REAL copied unchanged; empty slot search returns smallest index in 1..10.
*)
(* CONTRACT_RULES [] *)

recipeAdded := FALSE;
recipeDeleted := FALSE;
recipeModified := FALSE;
error := FALSE;
status := 0;
recipeQueryResult := tmp_blankRecipe;
tmp_commandCount := 0;
tmp_foundIndex := 0;
tmp_emptyIndex := 0;
tmp_duplicateFound := FALSE;

IF addRecipe THEN
    tmp_commandCount := tmp_commandCount + 1;
END_IF;
IF deleteRecipe THEN
    tmp_commandCount := tmp_commandCount + 1;
END_IF;
IF modifyRecipe THEN
    tmp_commandCount := tmp_commandCount + 1;
END_IF;
IF queryRecipe THEN
    tmp_commandCount := tmp_commandCount + 1;
END_IF;

IF tmp_commandCount > 1 THEN
    error := TRUE;
    status := 16#8000;

ELSIF addRecipe THEN
    FOR tmp_i := 1 TO 10 DO
        IF (recipe[tmp_i].recipeID <> 0) AND (recipe[tmp_i].recipeID = recipeIn.recipeID) THEN
            tmp_duplicateFound := TRUE;
        END_IF;
    END_FOR;

    IF tmp_duplicateFound THEN
        error := TRUE;
        status := 16#8002;
    ELSE
        FOR tmp_i := 1 TO 10 DO
            IF (recipe[tmp_i].recipeID = 0) AND (tmp_emptyIndex = 0) THEN
                tmp_emptyIndex := tmp_i;
            END_IF;
        END_FOR;

        IF tmp_emptyIndex = 0 THEN
            error := TRUE;
            status := 16#8003;
        ELSE
            recipe[tmp_emptyIndex] := recipeIn;
            recipeAdded := TRUE;
        END_IF;
    END_IF;

ELSIF deleteRecipe THEN
    FOR tmp_i := 1 TO 10 DO
        IF (recipe[tmp_i].recipeID <> 0) AND (recipe[tmp_i].recipeID = recipeIn.recipeID) THEN
            tmp_foundIndex := tmp_i;
        END_IF;
    END_FOR;

    IF tmp_foundIndex = 0 THEN
        error := TRUE;
        status := 16#8004;
    ELSE
        recipe[tmp_foundIndex].recipeID := 0;
        recipeDeleted := TRUE;
    END_IF;

ELSIF modifyRecipe THEN
    FOR tmp_i := 1 TO 10 DO
        IF (recipe[tmp_i].recipeID <> 0) AND (recipe[tmp_i].recipeID = recipeIn.recipeID) THEN
            tmp_foundIndex := tmp_i;
        END_IF;
    END_FOR;

    IF tmp_foundIndex = 0 THEN
        error := TRUE;
        status := 16#8005;
    ELSE
        recipe[tmp_foundIndex] := recipeIn;
        recipeModified := TRUE;
    END_IF;

ELSIF queryRecipe THEN
    FOR tmp_i := 1 TO 10 DO
        IF (recipe[tmp_i].recipeID <> 0) AND (recipe[tmp_i].recipeID = recipeIn.recipeID) THEN
            tmp_foundIndex := tmp_i;
        END_IF;
    END_FOR;

    IF tmp_foundIndex = 0 THEN
        error := TRUE;
        status := 16#8001;
    ELSE
        recipeQueryResult := recipe[tmp_foundIndex];
    END_IF;
END_IF;

(* ---- public-hard-03.candidate_02.st ---- *)
TYPE ST_Recipe :
STRUCT
    recipeID : INT;
    ingredientType : INT;
    ingredientRatio : REAL;
    productionTemperature : REAL;
END_STRUCT
END_TYPE;

FUNCTION_BLOCK FB_RecipeManagementSystem
VAR_INPUT
    addRecipe : BOOL;
    deleteRecipe : BOOL;
    modifyRecipe : BOOL;
    queryRecipe : BOOL;
    recipeIn : ST_Recipe;
END_VAR
VAR_OUTPUT
    recipeAdded : BOOL;
    recipeDeleted : BOOL;
    recipeModified : BOOL;
    recipeQueryResult : ST_Recipe;
    error : BOOL;
    status : WORD;
END_VAR
VAR_IN_OUT
    recipe : ARRAY[1..10] OF ST_Recipe;
END_VAR
VAR
    tmp_i : INT;
    tmp_foundIndex : INT;
    tmp_emptyIndex : INT;
    tmp_duplicateFound : BOOL;
    tmp_commandCount : INT;
    tmp_blankRecipe : ST_Recipe;
END_VAR

(* ENGINEERING_CONTRACT
   recipeAdded/Deleted/Modified: pulse TRUE only in the scan of a successful sole command; no retention; cleared each scan.
   recipeQueryResult: assigned from the matched recipe on a successful sole query; cleared to blank on all other scans; no retention.
   error/status: combinational per scan; PUB002-PUB006 error codes 16#8001..16#8005 on sole-command failures; 16#0000 on success/no operation.
   database recipe: retained through IN_OUT; altered only by successful add/delete/modify per PUB003-PUB005; slot recipeID=0 means empty.
   same-scan priority: simultaneous command requests are reported as unsupported with 16#8000; PUB011 leaves this case unspecified.
   units/boundaries: identifiers INT, ratios/temperatures REAL copied unchanged; empty slot search returns smallest index in 1..10.
*)
(* CONTRACT_RULES [] *)

recipeAdded := FALSE;
recipeDeleted := FALSE;
recipeModified := FALSE;
error := FALSE;
status := 0;
recipeQueryResult := tmp_blankRecipe;
tmp_commandCount := 0;
tmp_foundIndex := 0;
tmp_emptyIndex := 0;
tmp_duplicateFound := FALSE;

IF addRecipe THEN
    tmp_commandCount := tmp_commandCount + 1;
END_IF;
IF deleteRecipe THEN
    tmp_commandCount := tmp_commandCount + 1;
END_IF;
IF modifyRecipe THEN
    tmp_commandCount := tmp_commandCount + 1;
END_IF;
IF queryRecipe THEN
    tmp_commandCount := tmp_commandCount + 1;
END_IF;

IF tmp_commandCount > 1 THEN
    error := TRUE;
    status := 16#8000;

ELSIF addRecipe THEN
    FOR tmp_i := 1 TO 10 DO
        IF (recipe[tmp_i].recipeID <> 0) AND (recipe[tmp_i].recipeID = recipeIn.recipeID) THEN
            tmp_duplicateFound := TRUE;
        END_IF;
    END_FOR;

    IF tmp_duplicateFound THEN
        error := TRUE;
        status := 16#8002;
    ELSE
        FOR tmp_i := 1 TO 10 DO
            IF (recipe[tmp_i].recipeID = 0) AND (tmp_emptyIndex = 0) THEN
                tmp_emptyIndex := tmp_i;
            END_IF;
        END_FOR;

        IF tmp_emptyIndex = 0 THEN
            error := TRUE;
            status := 16#8003;
        ELSE
            recipe[tmp_emptyIndex] := recipeIn;
            recipeAdded := TRUE;
        END_IF;
    END_IF;

ELSIF deleteRecipe THEN
    FOR tmp_i := 1 TO 10 DO
        IF (recipe[tmp_i].recipeID <> 0) AND (recipe[tmp_i].recipeID = recipeIn.recipeID) THEN
            tmp_foundIndex := tmp_i;
        END_IF;
    END_FOR;

    IF tmp_foundIndex = 0 THEN
        error := TRUE;
        status := 16#8004;
    ELSE
        recipe[tmp_foundIndex].recipeID := 0;
        recipeDeleted := TRUE;
    END_IF;

ELSIF modifyRecipe THEN
    FOR tmp_i := 1 TO 10 DO
        IF (recipe[tmp_i].recipeID <> 0) AND (recipe[tmp_i].recipeID = recipeIn.recipeID) THEN
            tmp_foundIndex := tmp_i;
        END_IF;
    END_FOR;

    IF tmp_foundIndex = 0 THEN
        error := TRUE;
        status := 16#8005;
    ELSE
        recipe[tmp_foundIndex] := recipeIn;
        recipeModified := TRUE;
    END_IF;

ELSIF queryRecipe THEN
    FOR tmp_i := 1 TO 10 DO
        IF (recipe[tmp_i].recipeID <> 0) AND (recipe[tmp_i].recipeID = recipeIn.recipeID) THEN
            tmp_foundIndex := tmp_i;
        END_IF;
    END_FOR;

    IF tmp_foundIndex = 0 THEN
        error := TRUE;
        status := 16#8001;
    ELSE
        recipeQueryResult := recipe[tmp_foundIndex];
    END_IF;
END_IF;

END_FUNCTION_BLOCK

(* ---- public-hard-03.candidate_03.st ---- *)
TYPE ST_Recipe :
STRUCT
    recipeID : INT;
    ingredientType : INT;
    ingredientRatio : REAL;
    productionTemperature : REAL;
END_STRUCT
END_TYPE;

FUNCTION_BLOCK FB_RecipeManagementSystem
VAR_INPUT
    addRecipe : BOOL;
    deleteRecipe : BOOL;
    modifyRecipe : BOOL;
    queryRecipe : BOOL;
    recipeIn : ST_Recipe;
END_VAR
VAR_OUTPUT
    recipeAdded : BOOL;
    recipeDeleted : BOOL;
    recipeModified : BOOL;
    recipeQueryResult : ST_Recipe;
    error : BOOL;
    status : WORD;
END_VAR
VAR_IN_OUT
    recipe : ARRAY[1..10] OF ST_Recipe;
END_VAR
VAR
    tmp_i : INT;
    tmp_foundIndex : INT;
    tmp_emptyIndex : INT;
    tmp_duplicateFound : BOOL;
    tmp_commandCount : INT;

END_VAR

(* ENGINEERING_CONTRACT
   recipeAdded/Deleted/Modified: pulse TRUE only in the scan of a successful sole command; no retention; cleared each scan.
   recipeQueryResult: assigned from the matched recipe on a successful sole query; retains its last value otherwise.
   error/status: combinational per scan; PUB002-PUB006 error codes 16#8001..16#8005 on sole-command failures; 16#0000 on success/no operation.
   database recipe: retained through IN_OUT; altered only by successful add/delete/modify per PUB003-PUB005; slot recipeID=0 means empty.
   same-scan priority: simultaneous command requests are reported as unsupported with 16#8000; PUB011 leaves this case unspecified.
   units/boundaries: identifiers INT, ratios/temperatures REAL copied unchanged; empty slot search returns smallest index in 1..10.
*)
(* CONTRACT_RULES [] *)

recipeAdded := FALSE;
recipeDeleted := FALSE;
recipeModified := FALSE;
error := FALSE;
status := 0;

tmp_commandCount := 0;
tmp_foundIndex := 0;
tmp_emptyIndex := 0;
tmp_duplicateFound := FALSE;

IF addRecipe THEN
    tmp_commandCount := tmp_commandCount + 1;
END_IF;
IF deleteRecipe THEN
    tmp_commandCount := tmp_commandCount + 1;
END_IF;
IF modifyRecipe THEN
    tmp_commandCount := tmp_commandCount + 1;
END_IF;
IF queryRecipe THEN
    tmp_commandCount := tmp_commandCount + 1;
END_IF;

IF tmp_commandCount > 1 THEN
    error := TRUE;
    status := 16#8000;

ELSIF addRecipe THEN
    FOR tmp_i := 1 TO 10 DO
        IF (recipe[tmp_i].recipeID <> 0) AND (recipe[tmp_i].recipeID = recipeIn.recipeID) THEN
            tmp_duplicateFound := TRUE;
        END_IF;
    END_FOR;

    IF tmp_duplicateFound THEN
        error := TRUE;
        status := 16#8002;
    ELSE
        FOR tmp_i := 1 TO 10 DO
            IF (recipe[tmp_i].recipeID = 0) AND (tmp_emptyIndex = 0) THEN
                tmp_emptyIndex := tmp_i;
            END_IF;
        END_FOR;

        IF tmp_emptyIndex = 0 THEN
            error := TRUE;
            status := 16#8003;
        ELSE
            recipe[tmp_emptyIndex] := recipeIn;
            recipeAdded := TRUE;
        END_IF;
    END_IF;

ELSIF deleteRecipe THEN
    FOR tmp_i := 1 TO 10 DO
        IF (recipe[tmp_i].recipeID <> 0) AND (recipe[tmp_i].recipeID = recipeIn.recipeID) THEN
            tmp_foundIndex := tmp_i;
        END_IF;
    END_FOR;

    IF tmp_foundIndex = 0 THEN
        error := TRUE;
        status := 16#8004;
    ELSE
        recipe[tmp_foundIndex].recipeID := 0;
        recipeDeleted := TRUE;
    END_IF;

ELSIF modifyRecipe THEN
    FOR tmp_i := 1 TO 10 DO
        IF (recipe[tmp_i].recipeID <> 0) AND (recipe[tmp_i].recipeID = recipeIn.recipeID) THEN
            tmp_foundIndex := tmp_i;
        END_IF;
    END_FOR;

    IF tmp_foundIndex = 0 THEN
        error := TRUE;
        status := 16#8005;
    ELSE
        recipe[tmp_foundIndex] := recipeIn;
        recipeModified := TRUE;
    END_IF;

ELSIF queryRecipe THEN
    FOR tmp_i := 1 TO 10 DO
        IF (recipe[tmp_i].recipeID <> 0) AND (recipe[tmp_i].recipeID = recipeIn.recipeID) THEN
            tmp_foundIndex := tmp_i;
        END_IF;
    END_FOR;

    IF tmp_foundIndex = 0 THEN
        error := TRUE;
        status := 16#8001;
    ELSE
        recipeQueryResult := recipe[tmp_foundIndex];
    END_IF;
END_IF;

END_FUNCTION_BLOCK

(* ---- public-hard-03.patch_base_02.st ---- *)
TYPE ST_Recipe :
STRUCT
    recipeID : INT;
    ingredientType : INT;
    ingredientRatio : REAL;
    productionTemperature : REAL;
END_STRUCT
END_TYPE;

FUNCTION_BLOCK FB_RecipeManagementSystem
VAR_INPUT
    addRecipe : BOOL;
    deleteRecipe : BOOL;
    modifyRecipe : BOOL;
    queryRecipe : BOOL;
    recipeIn : ST_Recipe;
END_VAR
VAR_OUTPUT
    recipeAdded : BOOL;
    recipeDeleted : BOOL;
    recipeModified : BOOL;
    recipeQueryResult : ST_Recipe;
    error : BOOL;
    status : WORD;
END_VAR
VAR_IN_OUT
    recipe : ARRAY[1..10] OF ST_Recipe;
END_VAR
VAR
    tmp_i : INT;
    tmp_foundIndex : INT;
    tmp_emptyIndex : INT;
    tmp_duplicateFound : BOOL;
    tmp_commandCount : INT;
    tmp_blankRecipe : ST_Recipe;
END_VAR

(* ENGINEERING_CONTRACT
   recipeAdded/Deleted/Modified: pulse TRUE only in the scan of a successful sole command; no retention; cleared each scan.
   recipeQueryResult: assigned from the matched recipe on a successful sole query; cleared to blank on all other scans; no retention.
   error/status: combinational per scan; PUB002-PUB006 error codes 16#8001..16#8005 on sole-command failures; 16#0000 on success/no operation.
   database recipe: retained through IN_OUT; altered only by successful add/delete/modify per PUB003-PUB005; slot recipeID=0 means empty.
   same-scan priority: simultaneous command requests are reported as unsupported with 16#8000; PUB011 leaves this case unspecified.
   units/boundaries: identifiers INT, ratios/temperatures REAL copied unchanged; empty slot search returns smallest index in 1..10.
*)
(* CONTRACT_RULES [] *)

recipeAdded := FALSE;
recipeDeleted := FALSE;
recipeModified := FALSE;
error := FALSE;
status := 0;
recipeQueryResult := tmp_blankRecipe;
tmp_commandCount := 0;
tmp_foundIndex := 0;
tmp_emptyIndex := 0;
tmp_duplicateFound := FALSE;

IF addRecipe THEN
    tmp_commandCount := tmp_commandCount + 1;
END_IF;
IF deleteRecipe THEN
    tmp_commandCount := tmp_commandCount + 1;
END_IF;
IF modifyRecipe THEN
    tmp_commandCount := tmp_commandCount + 1;
END_IF;
IF queryRecipe THEN
    tmp_commandCount := tmp_commandCount + 1;
END_IF;

IF tmp_commandCount > 1 THEN
    error := TRUE;
    status := 16#8000;

ELSIF addRecipe THEN
    FOR tmp_i := 1 TO 10 DO
        IF (recipe[tmp_i].recipeID <> 0) AND (recipe[tmp_i].recipeID = recipeIn.recipeID) THEN
            tmp_duplicateFound := TRUE;
        END_IF;
    END_FOR;

    IF tmp_duplicateFound THEN
        error := TRUE;
        status := 16#8002;
    ELSE
        FOR tmp_i := 1 TO 10 DO
            IF (recipe[tmp_i].recipeID = 0) AND (tmp_emptyIndex = 0) THEN
                tmp_emptyIndex := tmp_i;
            END_IF;
        END_FOR;

        IF tmp_emptyIndex = 0 THEN
            error := TRUE;
            status := 16#8003;
        ELSE
            recipe[tmp_emptyIndex] := recipeIn;
            recipeAdded := TRUE;
        END_IF;
    END_IF;

ELSIF deleteRecipe THEN
    FOR tmp_i := 1 TO 10 DO
        IF (recipe[tmp_i].recipeID <> 0) AND (recipe[tmp_i].recipeID = recipeIn.recipeID) THEN
            tmp_foundIndex := tmp_i;
        END_IF;
    END_FOR;

    IF tmp_foundIndex = 0 THEN
        error := TRUE;
        status := 16#8004;
    ELSE
        recipe[tmp_foundIndex].recipeID := 0;
        recipeDeleted := TRUE;
    END_IF;

ELSIF modifyRecipe THEN
    FOR tmp_i := 1 TO 10 DO
        IF (recipe[tmp_i].recipeID <> 0) AND (recipe[tmp_i].recipeID = recipeIn.recipeID) THEN
            tmp_foundIndex := tmp_i;
        END_IF;
    END_FOR;

    IF tmp_foundIndex = 0 THEN
        error := TRUE;
        status := 16#8005;
    ELSE
        recipe[tmp_foundIndex] := recipeIn;
        recipeModified := TRUE;
    END_IF;

ELSIF queryRecipe THEN
    FOR tmp_i := 1 TO 10 DO
        IF (recipe[tmp_i].recipeID <> 0) AND (recipe[tmp_i].recipeID = recipeIn.recipeID) THEN
            tmp_foundIndex := tmp_i;
        END_IF;
    END_FOR;

    IF tmp_foundIndex = 0 THEN
        error := TRUE;
        status := 16#8001;
    ELSE
        recipeQueryResult := recipe[tmp_foundIndex];
    END_IF;
END_IF;

(* ---- public-hard-03.patch_base_03.st ---- *)
TYPE ST_Recipe :
STRUCT
    recipeID : INT;
    ingredientType : INT;
    ingredientRatio : REAL;
    productionTemperature : REAL;
END_STRUCT
END_TYPE;

FUNCTION_BLOCK FB_RecipeManagementSystem
VAR_INPUT
    addRecipe : BOOL;
    deleteRecipe : BOOL;
    modifyRecipe : BOOL;
    queryRecipe : BOOL;
    recipeIn : ST_Recipe;
END_VAR
VAR_OUTPUT
    recipeAdded : BOOL;
    recipeDeleted : BOOL;
    recipeModified : BOOL;
    recipeQueryResult : ST_Recipe;
    error : BOOL;
    status : WORD;
END_VAR
VAR_IN_OUT
    recipe : ARRAY[1..10] OF ST_Recipe;
END_VAR
VAR
    tmp_i : INT;
    tmp_foundIndex : INT;
    tmp_emptyIndex : INT;
    tmp_duplicateFound : BOOL;
    tmp_commandCount : INT;
    tmp_blankRecipe : ST_Recipe;
END_VAR

(* ENGINEERING_CONTRACT
   recipeAdded/Deleted/Modified: pulse TRUE only in the scan of a successful sole command; no retention; cleared each scan.
   recipeQueryResult: assigned from the matched recipe on a successful sole query; cleared to blank on all other scans; no retention.
   error/status: combinational per scan; PUB002-PUB006 error codes 16#8001..16#8005 on sole-command failures; 16#0000 on success/no operation.
   database recipe: retained through IN_OUT; altered only by successful add/delete/modify per PUB003-PUB005; slot recipeID=0 means empty.
   same-scan priority: simultaneous command requests are reported as unsupported with 16#8000; PUB011 leaves this case unspecified.
   units/boundaries: identifiers INT, ratios/temperatures REAL copied unchanged; empty slot search returns smallest index in 1..10.
*)
(* CONTRACT_RULES [] *)

recipeAdded := FALSE;
recipeDeleted := FALSE;
recipeModified := FALSE;
error := FALSE;
status := 0;
recipeQueryResult := tmp_blankRecipe;
tmp_commandCount := 0;
tmp_foundIndex := 0;
tmp_emptyIndex := 0;
tmp_duplicateFound := FALSE;

IF addRecipe THEN
    tmp_commandCount := tmp_commandCount + 1;
END_IF;
IF deleteRecipe THEN
    tmp_commandCount := tmp_commandCount + 1;
END_IF;
IF modifyRecipe THEN
    tmp_commandCount := tmp_commandCount + 1;
END_IF;
IF queryRecipe THEN
    tmp_commandCount := tmp_commandCount + 1;
END_IF;

IF tmp_commandCount > 1 THEN
    error := TRUE;
    status := 16#8000;

ELSIF addRecipe THEN
    FOR tmp_i := 1 TO 10 DO
        IF (recipe[tmp_i].recipeID <> 0) AND (recipe[tmp_i].recipeID = recipeIn.recipeID) THEN
            tmp_duplicateFound := TRUE;
        END_IF;
    END_FOR;

    IF tmp_duplicateFound THEN
        error := TRUE;
        status := 16#8002;
    ELSE
        FOR tmp_i := 1 TO 10 DO
            IF (recipe[tmp_i].recipeID = 0) AND (tmp_emptyIndex = 0) THEN
                tmp_emptyIndex := tmp_i;
            END_IF;
        END_FOR;

        IF tmp_emptyIndex = 0 THEN
            error := TRUE;
            status := 16#8003;
        ELSE
            recipe[tmp_emptyIndex] := recipeIn;
            recipeAdded := TRUE;
        END_IF;
    END_IF;

ELSIF deleteRecipe THEN
    FOR tmp_i := 1 TO 10 DO
        IF (recipe[tmp_i].recipeID <> 0) AND (recipe[tmp_i].recipeID = recipeIn.recipeID) THEN
            tmp_foundIndex := tmp_i;
        END_IF;
    END_FOR;

    IF tmp_foundIndex = 0 THEN
        error := TRUE;
        status := 16#8004;
    ELSE
        recipe[tmp_foundIndex].recipeID := 0;
        recipeDeleted := TRUE;
    END_IF;

ELSIF modifyRecipe THEN
    FOR tmp_i := 1 TO 10 DO
        IF (recipe[tmp_i].recipeID <> 0) AND (recipe[tmp_i].recipeID = recipeIn.recipeID) THEN
            tmp_foundIndex := tmp_i;
        END_IF;
    END_FOR;

    IF tmp_foundIndex = 0 THEN
        error := TRUE;
        status := 16#8005;
    ELSE
        recipe[tmp_foundIndex] := recipeIn;
        recipeModified := TRUE;
    END_IF;

ELSIF queryRecipe THEN
    FOR tmp_i := 1 TO 10 DO
        IF (recipe[tmp_i].recipeID <> 0) AND (recipe[tmp_i].recipeID = recipeIn.recipeID) THEN
            tmp_foundIndex := tmp_i;
        END_IF;
    END_FOR;

    IF tmp_foundIndex = 0 THEN
        error := TRUE;
        status := 16#8001;
    ELSE
        recipeQueryResult := recipe[tmp_foundIndex];
    END_IF;
END_IF;

END_FUNCTION_BLOCK

(* ---- public-hard-03.raw_candidate_01.st ---- *)
TYPE ST_Recipe :
STRUCT
    recipeID : INT;
    ingredientType : INT;
    ingredientRatio : REAL;
    productionTemperature : REAL;
END_STRUCT
END_TYPE

FUNCTION_BLOCK FB_RecipeManagementSystem
VAR_INPUT
    addRecipe : BOOL;
    deleteRecipe : BOOL;
    modifyRecipe : BOOL;
    queryRecipe : BOOL;
    recipeIn : ST_Recipe;
END_VAR
VAR_OUTPUT
    recipeAdded : BOOL;
    recipeDeleted : BOOL;
    recipeModified : BOOL;
    recipeQueryResult : ST_Recipe;
    error : BOOL;
    status : WORD;
END_VAR
VAR_IN_OUT
    recipe : ARRAY[1..10] OF ST_Recipe;
END_VAR
VAR
    tmp_i : INT;
    tmp_foundIndex : INT;
    tmp_emptyIndex : INT;
    tmp_duplicateFound : BOOL;
    tmp_commandCount : INT;
    tmp_blankRecipe : ST_Recipe;
END_VAR

(* ENGINEERING_CONTRACT
   recipeAdded/Deleted/Modified: pulse TRUE only in the scan of a successful sole command; no retention; cleared each scan.
   recipeQueryResult: assigned from the matched recipe on a successful sole query; cleared to blank on all other scans; no retention.
   error/status: combinational per scan; PUB002-PUB006 error codes 16#8001..16#8005 on sole-command failures; 16#0000 on success/no operation.
   database recipe: retained through IN_OUT; altered only by successful add/delete/modify per PUB003-PUB005; slot recipeID=0 means empty.
   same-scan priority: simultaneous command requests are reported as unsupported with 16#8000; PUB011 leaves this case unspecified.
   units/boundaries: identifiers INT, ratios/temperatures REAL copied unchanged; empty slot search returns smallest index in 1..10.
*)
(* CONTRACT_RULES [] *)

recipeAdded := FALSE;
recipeDeleted := FALSE;
recipeModified := FALSE;
error := FALSE;
status := 0;
recipeQueryResult := tmp_blankRecipe;
tmp_commandCount := 0;
tmp_foundIndex := 0;
tmp_emptyIndex := 0;
tmp_duplicateFound := FALSE;

IF addRecipe THEN
    tmp_commandCount := tmp_commandCount + 1;
END_IF;
IF deleteRecipe THEN
    tmp_commandCount := tmp_commandCount + 1;
END_IF;
IF modifyRecipe THEN
    tmp_commandCount := tmp_commandCount + 1;
END_IF;
IF queryRecipe THEN
    tmp_commandCount := tmp_commandCount + 1;
END_IF;

IF tmp_commandCount > 1 THEN
    error := TRUE;
    status := 16#8000;

ELSIF addRecipe THEN
    FOR tmp_i := 1 TO 10 DO
        IF (recipe[tmp_i].recipeID <> 0) AND (recipe[tmp_i].recipeID = recipeIn.recipeID) THEN
            tmp_duplicateFound := TRUE;
        END_IF;
    END_FOR;

    IF tmp_duplicateFound THEN
        error := TRUE;
        status := 16#8002;
    ELSE
        FOR tmp_i := 1 TO 10 DO
            IF (recipe[tmp_i].recipeID = 0) AND (tmp_emptyIndex = 0) THEN
                tmp_emptyIndex := tmp_i;
            END_IF;
        END_FOR;

        IF tmp_emptyIndex = 0 THEN
            error := TRUE;
            status := 16#8003;
        ELSE
            recipe[tmp_emptyIndex] := recipeIn;
            recipeAdded := TRUE;
        END_IF;
    END_IF;

ELSIF deleteRecipe THEN
    FOR tmp_i := 1 TO 10 DO
        IF (recipe[tmp_i].recipeID <> 0) AND (recipe[tmp_i].recipeID = recipeIn.recipeID) THEN
            tmp_foundIndex := tmp_i;
        END_IF;
    END_FOR;

    IF tmp_foundIndex = 0 THEN
        error := TRUE;
        status := 16#8004;
    ELSE
        recipe[tmp_foundIndex].recipeID := 0;
        recipeDeleted := TRUE;
    END_IF;

ELSIF modifyRecipe THEN
    FOR tmp_i := 1 TO 10 DO
        IF (recipe[tmp_i].recipeID <> 0) AND (recipe[tmp_i].recipeID = recipeIn.recipeID) THEN
            tmp_foundIndex := tmp_i;
        END_IF;
    END_FOR;

    IF tmp_foundIndex = 0 THEN
        error := TRUE;
        status := 16#8005;
    ELSE
        recipe[tmp_foundIndex] := recipeIn;
        recipeModified := TRUE;
    END_IF;

ELSIF queryRecipe THEN
    FOR tmp_i := 1 TO 10 DO
        IF (recipe[tmp_i].recipeID <> 0) AND (recipe[tmp_i].recipeID = recipeIn.recipeID) THEN
            tmp_foundIndex := tmp_i;
        END_IF;
    END_FOR;

    IF tmp_foundIndex = 0 THEN
        error := TRUE;
        status := 16#8001;
    ELSE
        recipeQueryResult := recipe[tmp_foundIndex];
    END_IF;
END_IF;

(* ---- public-hard-03.raw_candidate_02.st ---- *)
TYPE ST_Recipe :
STRUCT
    recipeID : INT;
    ingredientType : INT;
    ingredientRatio : REAL;
    productionTemperature : REAL;
END_STRUCT
END_TYPE;

FUNCTION_BLOCK FB_RecipeManagementSystem
VAR_INPUT
    addRecipe : BOOL;
    deleteRecipe : BOOL;
    modifyRecipe : BOOL;
    queryRecipe : BOOL;
    recipeIn : ST_Recipe;
END_VAR
VAR_OUTPUT
    recipeAdded : BOOL;
    recipeDeleted : BOOL;
    recipeModified : BOOL;
    recipeQueryResult : ST_Recipe;
    error : BOOL;
    status : WORD;
END_VAR
VAR_IN_OUT
    recipe : ARRAY[1..10] OF ST_Recipe;
END_VAR
VAR
    tmp_i : INT;
    tmp_foundIndex : INT;
    tmp_emptyIndex : INT;
    tmp_duplicateFound : BOOL;
    tmp_commandCount : INT;
    tmp_blankRecipe : ST_Recipe;
END_VAR

(* ENGINEERING_CONTRACT
   recipeAdded/Deleted/Modified: pulse TRUE only in the scan of a successful sole command; no retention; cleared each scan.
   recipeQueryResult: assigned from the matched recipe on a successful sole query; cleared to blank on all other scans; no retention.
   error/status: combinational per scan; PUB002-PUB006 error codes 16#8001..16#8005 on sole-command failures; 16#0000 on success/no operation.
   database recipe: retained through IN_OUT; altered only by successful add/delete/modify per PUB003-PUB005; slot recipeID=0 means empty.
   same-scan priority: simultaneous command requests are reported as unsupported with 16#8000; PUB011 leaves this case unspecified.
   units/boundaries: identifiers INT, ratios/temperatures REAL copied unchanged; empty slot search returns smallest index in 1..10.
*)
(* CONTRACT_RULES [] *)

recipeAdded := FALSE;
recipeDeleted := FALSE;
recipeModified := FALSE;
error := FALSE;
status := 0;
recipeQueryResult := tmp_blankRecipe;
tmp_commandCount := 0;
tmp_foundIndex := 0;
tmp_emptyIndex := 0;
tmp_duplicateFound := FALSE;

IF addRecipe THEN
    tmp_commandCount := tmp_commandCount + 1;
END_IF;
IF deleteRecipe THEN
    tmp_commandCount := tmp_commandCount + 1;
END_IF;
IF modifyRecipe THEN
    tmp_commandCount := tmp_commandCount + 1;
END_IF;
IF queryRecipe THEN
    tmp_commandCount := tmp_commandCount + 1;
END_IF;

IF tmp_commandCount > 1 THEN
    error := TRUE;
    status := 16#8000;

ELSIF addRecipe THEN
    FOR tmp_i := 1 TO 10 DO
        IF (recipe[tmp_i].recipeID <> 0) AND (recipe[tmp_i].recipeID = recipeIn.recipeID) THEN
            tmp_duplicateFound := TRUE;
        END_IF;
    END_FOR;

    IF tmp_duplicateFound THEN
        error := TRUE;
        status := 16#8002;
    ELSE
        FOR tmp_i := 1 TO 10 DO
            IF (recipe[tmp_i].recipeID = 0) AND (tmp_emptyIndex = 0) THEN
                tmp_emptyIndex := tmp_i;
            END_IF;
        END_FOR;

        IF tmp_emptyIndex = 0 THEN
            error := TRUE;
            status := 16#8003;
        ELSE
            recipe[tmp_emptyIndex] := recipeIn;
            recipeAdded := TRUE;
        END_IF;
    END_IF;

ELSIF deleteRecipe THEN
    FOR tmp_i := 1 TO 10 DO
        IF (recipe[tmp_i].recipeID <> 0) AND (recipe[tmp_i].recipeID = recipeIn.recipeID) THEN
            tmp_foundIndex := tmp_i;
        END_IF;
    END_FOR;

    IF tmp_foundIndex = 0 THEN
        error := TRUE;
        status := 16#8004;
    ELSE
        recipe[tmp_foundIndex].recipeID := 0;
        recipeDeleted := TRUE;
    END_IF;

ELSIF modifyRecipe THEN
    FOR tmp_i := 1 TO 10 DO
        IF (recipe[tmp_i].recipeID <> 0) AND (recipe[tmp_i].recipeID = recipeIn.recipeID) THEN
            tmp_foundIndex := tmp_i;
        END_IF;
    END_FOR;

    IF tmp_foundIndex = 0 THEN
        error := TRUE;
        status := 16#8005;
    ELSE
        recipe[tmp_foundIndex] := recipeIn;
        recipeModified := TRUE;
    END_IF;

ELSIF queryRecipe THEN
    FOR tmp_i := 1 TO 10 DO
        IF (recipe[tmp_i].recipeID <> 0) AND (recipe[tmp_i].recipeID = recipeIn.recipeID) THEN
            tmp_foundIndex := tmp_i;
        END_IF;
    END_FOR;

    IF tmp_foundIndex = 0 THEN
        error := TRUE;
        status := 16#8001;
    ELSE
        recipeQueryResult := recipe[tmp_foundIndex];
    END_IF;
END_IF;

END_FUNCTION_BLOCK

(* ---- public-hard-03.raw_candidate_03.st ---- *)
TYPE ST_Recipe :
STRUCT
    recipeID : INT;
    ingredientType : INT;
    ingredientRatio : REAL;
    productionTemperature : REAL;
END_STRUCT
END_TYPE;

FUNCTION_BLOCK FB_RecipeManagementSystem
VAR_INPUT
    addRecipe : BOOL;
    deleteRecipe : BOOL;
    modifyRecipe : BOOL;
    queryRecipe : BOOL;
    recipeIn : ST_Recipe;
END_VAR
VAR_OUTPUT
    recipeAdded : BOOL;
    recipeDeleted : BOOL;
    recipeModified : BOOL;
    recipeQueryResult : ST_Recipe;
    error : BOOL;
    status : WORD;
END_VAR
VAR_IN_OUT
    recipe : ARRAY[1..10] OF ST_Recipe;
END_VAR
VAR
    tmp_i : INT;
    tmp_foundIndex : INT;
    tmp_emptyIndex : INT;
    tmp_duplicateFound : BOOL;
    tmp_commandCount : INT;

END_VAR

(* ENGINEERING_CONTRACT
   recipeAdded/Deleted/Modified: pulse TRUE only in the scan of a successful sole command; no retention; cleared each scan.
   recipeQueryResult: assigned from the matched recipe on a successful sole query; retains its last value otherwise.
   error/status: combinational per scan; PUB002-PUB006 error codes 16#8001..16#8005 on sole-command failures; 16#0000 on success/no operation.
   database recipe: retained through IN_OUT; altered only by successful add/delete/modify per PUB003-PUB005; slot recipeID=0 means empty.
   same-scan priority: simultaneous command requests are reported as unsupported with 16#8000; PUB011 leaves this case unspecified.
   units/boundaries: identifiers INT, ratios/temperatures REAL copied unchanged; empty slot search returns smallest index in 1..10.
*)
(* CONTRACT_RULES [] *)

recipeAdded := FALSE;
recipeDeleted := FALSE;
recipeModified := FALSE;
error := FALSE;
status := 0;

tmp_commandCount := 0;
tmp_foundIndex := 0;
tmp_emptyIndex := 0;
tmp_duplicateFound := FALSE;

IF addRecipe THEN
    tmp_commandCount := tmp_commandCount + 1;
END_IF;
IF deleteRecipe THEN
    tmp_commandCount := tmp_commandCount + 1;
END_IF;
IF modifyRecipe THEN
    tmp_commandCount := tmp_commandCount + 1;
END_IF;
IF queryRecipe THEN
    tmp_commandCount := tmp_commandCount + 1;
END_IF;

IF tmp_commandCount > 1 THEN
    error := TRUE;
    status := 16#8000;

ELSIF addRecipe THEN
    FOR tmp_i := 1 TO 10 DO
        IF (recipe[tmp_i].recipeID <> 0) AND (recipe[tmp_i].recipeID = recipeIn.recipeID) THEN
            tmp_duplicateFound := TRUE;
        END_IF;
    END_FOR;

    IF tmp_duplicateFound THEN
        error := TRUE;
        status := 16#8002;
    ELSE
        FOR tmp_i := 1 TO 10 DO
            IF (recipe[tmp_i].recipeID = 0) AND (tmp_emptyIndex = 0) THEN
                tmp_emptyIndex := tmp_i;
            END_IF;
        END_FOR;

        IF tmp_emptyIndex = 0 THEN
            error := TRUE;
            status := 16#8003;
        ELSE
            recipe[tmp_emptyIndex] := recipeIn;
            recipeAdded := TRUE;
        END_IF;
    END_IF;

ELSIF deleteRecipe THEN
    FOR tmp_i := 1 TO 10 DO
        IF (recipe[tmp_i].recipeID <> 0) AND (recipe[tmp_i].recipeID = recipeIn.recipeID) THEN
            tmp_foundIndex := tmp_i;
        END_IF;
    END_FOR;

    IF tmp_foundIndex = 0 THEN
        error := TRUE;
        status := 16#8004;
    ELSE
        recipe[tmp_foundIndex].recipeID := 0;
        recipeDeleted := TRUE;
    END_IF;

ELSIF modifyRecipe THEN
    FOR tmp_i := 1 TO 10 DO
        IF (recipe[tmp_i].recipeID <> 0) AND (recipe[tmp_i].recipeID = recipeIn.recipeID) THEN
            tmp_foundIndex := tmp_i;
        END_IF;
    END_FOR;

    IF tmp_foundIndex = 0 THEN
        error := TRUE;
        status := 16#8005;
    ELSE
        recipe[tmp_foundIndex] := recipeIn;
        recipeModified := TRUE;
    END_IF;

ELSIF queryRecipe THEN
    FOR tmp_i := 1 TO 10 DO
        IF (recipe[tmp_i].recipeID <> 0) AND (recipe[tmp_i].recipeID = recipeIn.recipeID) THEN
            tmp_foundIndex := tmp_i;
        END_IF;
    END_FOR;

    IF tmp_foundIndex = 0 THEN
        error := TRUE;
        status := 16#8001;
    ELSE
        recipeQueryResult := recipe[tmp_foundIndex];
    END_IF;
END_IF;

END_FUNCTION_BLOCK

(* ---- public-hard-04.candidate_01.st ---- *)
FUNCTION_BLOCK FB
VAR_INPUT
    enqueue : BOOL;
    dequeue : BOOL;
    reset : BOOL;
END_VAR
VAR_OUTPUT
    elementCount : DINT;
    status : WORD;
END_VAR
VAR_IN_OUT
    item : VARIANT;
    buffer : VARIANT;
END_VAR
VAR
    tmp_enq_rise : R_TRIG;
    tmp_deq_rise : R_TRIG;
    tmp_enq_edge : BOOL;
    tmp_deq_edge : BOOL;
    tmp_lower : DINT;
    tmp_upper : DINT;
    tmp_capacity : DINT;
    tmp_head : DINT;
    tmp_tail : DINT;
    tmp_initialized : BOOL := FALSE;
END_VAR

(* ENGINEERING_CONTRACT
- elementCount: initialized to 0 on first invocation; incremented only after successful enqueue; decremented only after successful dequeue; set to 0 by reset.
- enqueue: rising edge appends item at tail and advances tail while elementCount < capacity; on full queue rejects with 16#8002 and leaves item unchanged (PUB001,PUB004,PUB005,PUB009).
- dequeue: rising edge writes buffer[head] back to item and advances head while elementCount > 0; on empty queue rejects with 16#8001 and leaves item unchanged (PUB002,PUB004,PUB005,PUB008).
- reset: TRUE empties the queue, sets elementCount to 0, and resets head/tail; reset has priority over enqueue/dequeue (PUB003).
- capacity: stored on first invocation as UPPER_BOUND(buffer,1)-LOWER_BOUND(buffer,1)+1; full means count equals capacity (PUB004,PUB010).
- status: reset to 16#0000 each invocation; rejection codes override no-error status (PUB006,PUB008,PUB009).
- enqueue+dequeue in the same invocation is caller-forbidden; implementation processes enqueue before dequeue for a deterministic forbidden-input result (PUB002).
*)

(* CONTRACT_RULES [] *)

tmp_enq_rise(CLK := enqueue);
tmp_deq_rise(CLK := dequeue);
tmp_enq_edge := tmp_enq_rise.Q;
tmp_deq_edge := tmp_deq_rise.Q;

IF NOT tmp_initialized THEN
    tmp_lower := TO_DINT(LOWER_BOUND(buffer, 1));
    tmp_upper := TO_DINT(UPPER_BOUND(buffer, 1));
    tmp_capacity := tmp_upper - tmp_lower + 1;
    tmp_head := tmp_lower;
    tmp_tail := tmp_lower;
    elementCount := 0;
    tmp_initialized := TRUE;
END_IF;

status := 16#0000;

IF reset THEN
    elementCount := 0;
    tmp_head := tmp_lower;
    tmp_tail := tmp_lower;
ELSE
    IF tmp_enq_edge THEN
        IF elementCount >= tmp_capacity THEN
            status := 16#8002;
        ELSE
            buffer[tmp_tail] := item;
            elementCount := elementCount + 1;
            tmp_tail := tmp_tail + 1;
            IF tmp_tail > tmp_upper THEN
                tmp_tail := tmp_lower;
            END_IF;
        END_IF;
    END_IF;

    IF tmp_deq_edge THEN
        IF elementCount <= 0 THEN
            status := 16#8001;
        ELSE
            item := buffer[tmp_head];
            elementCount := elementCount - 1;
            tmp_head := tmp_head + 1;
            IF tmp_head > tmp_upper THEN
                tmp_head := tmp_lower;
            END_IF;
        END_IF;
    END_IF;
END_IF;

END_FUNCTION_BLOCK

(* ---- public-hard-04.raw_candidate_01.st ---- *)
FUNCTION_BLOCK FB
VAR_INPUT
    enqueue : BOOL;
    dequeue : BOOL;
    reset : BOOL;
END_VAR
VAR_OUTPUT
    elementCount : DINT;
    status : WORD;
END_VAR
VAR_IN_OUT
    item : VARIANT;
    buffer : VARIANT;
END_VAR
VAR
    tmp_enq_rise : R_TRIG;
    tmp_deq_rise : R_TRIG;
    tmp_enq_edge : BOOL;
    tmp_deq_edge : BOOL;
    tmp_lower : DINT;
    tmp_upper : DINT;
    tmp_capacity : DINT;
    tmp_head : DINT;
    tmp_tail : DINT;
    tmp_initialized : BOOL := FALSE;
END_VAR

(* ENGINEERING_CONTRACT
- elementCount: initialized to 0 on first invocation; incremented only after successful enqueue; decremented only after successful dequeue; set to 0 by reset.
- enqueue: rising edge appends item at tail and advances tail while elementCount < capacity; on full queue rejects with 16#8002 and leaves item unchanged (PUB001,PUB004,PUB005,PUB009).
- dequeue: rising edge writes buffer[head] back to item and advances head while elementCount > 0; on empty queue rejects with 16#8001 and leaves item unchanged (PUB002,PUB004,PUB005,PUB008).
- reset: TRUE empties the queue, sets elementCount to 0, and resets head/tail; reset has priority over enqueue/dequeue (PUB003).
- capacity: stored on first invocation as UPPER_BOUND(buffer,1)-LOWER_BOUND(buffer,1)+1; full means count equals capacity (PUB004,PUB010).
- status: reset to 16#0000 each invocation; rejection codes override no-error status (PUB006,PUB008,PUB009).
- enqueue+dequeue in the same invocation is caller-forbidden; implementation processes enqueue before dequeue for a deterministic forbidden-input result (PUB002).
*)

(* CONTRACT_RULES [] *)

tmp_enq_rise(CLK := enqueue);
tmp_deq_rise(CLK := dequeue);
tmp_enq_edge := tmp_enq_rise.Q;
tmp_deq_edge := tmp_deq_rise.Q;

IF NOT tmp_initialized THEN
    tmp_lower := TO_DINT(LOWER_BOUND(buffer, 1));
    tmp_upper := TO_DINT(UPPER_BOUND(buffer, 1));
    tmp_capacity := tmp_upper - tmp_lower + 1;
    tmp_head := tmp_lower;
    tmp_tail := tmp_lower;
    elementCount := 0;
    tmp_initialized := TRUE;
END_IF;

status := 16#0000;

IF reset THEN
    elementCount := 0;
    tmp_head := tmp_lower;
    tmp_tail := tmp_lower;
ELSE
    IF tmp_enq_edge THEN
        IF elementCount >= tmp_capacity THEN
            status := 16#8002;
        ELSE
            buffer[tmp_tail] := item;
            elementCount := elementCount + 1;
            tmp_tail := tmp_tail + 1;
            IF tmp_tail > tmp_upper THEN
                tmp_tail := tmp_lower;
            END_IF;
        END_IF;
    END_IF;

    IF tmp_deq_edge THEN
        IF elementCount <= 0 THEN
            status := 16#8001;
        ELSE
            item := buffer[tmp_head];
            elementCount := elementCount - 1;
            tmp_head := tmp_head + 1;
            IF tmp_head > tmp_upper THEN
                tmp_head := tmp_lower;
            END_IF;
        END_IF;
    END_IF;
END_IF;

END_FUNCTION_BLOCK

(* ---- public-hard-05.candidate_01.st ---- *)
(* ENGINEERING_CONTRACT
   Manual axis output: ON while its button=1, opposite command inactive, and its limit=0; OFF on release/limit (PUB001).
   Manual grip/release: ON while button=1, opposite inactive, and its limit=0; OFF on release/limit (PUB001).
   Single-step: Start edge activates next index 0..7/wraps; output held until switch; next Start advances (PUB002-PUB003).
   Single-cycle: Start edge runs 0..7; holds each output until completion; stops after left; next Start restarts (PUB004).
   Continuous: Start edge runs 0..7 and loops after left while mode selected (PUB005).
   Emergency: EmergencyStop=FALSE overrides all outputs and freezes start/progression; state is retained (PUB006).
   Index completion: 0/4 DownLimit, 1 GripLimit, 2/6 UpLimit, 3 RightLimit, 5 ReleaseLimit, 7 LeftLimit.
   Same-scan priority: E-stop highest; a feedback-completed action cannot energize on its completion scan; next action starts next scan.
   Unspecified: post-E-stop resumption uses retained state; mode changes outside a mode retain sequence state.
*)
(* CONTRACT_RULES [] *)

FUNCTION_BLOCK MechanicalArmControl
VAR_INPUT
    ManualMode : BOOL;
    SingleStepMode : BOOL;
    SingleCycleMode : BOOL;
    ContinuousMode : BOOL;
    EmergencyStop : BOOL;
    Start : BOOL;
    DownButton : BOOL;
    UpButton : BOOL;
    LeftButton : BOOL;
    RightButton : BOOL;
    GripButton : BOOL;
    ReleaseButton : BOOL;
    DownLimitSwitch : BOOL;
    UpLimitSwitch : BOOL;
    LeftLimitSwitch : BOOL;
    RightLimitSwitch : BOOL;
    GripLimitSwitch : BOOL;
    ReleaseLimitSwitch : BOOL;
END_VAR
VAR_OUTPUT
    MoveDown : BOOL;
    MoveUp : BOOL;
    MoveLeft : BOOL;
    MoveRight : BOOL;
    ActivateGrip : BOOL;
    ActivateRelease : BOOL;
END_VAR
VAR
    tmp_startEdge : R_TRIG;
    tmp_autoMode : BOOL;
    tmp_autoActive : BOOL := FALSE;
    tmp_currentStep : INT := 0;
    tmp_singleNextStep : INT := 0;
    tmp_targetReached : BOOL;

    tmp_manualDownReq : BOOL;
    tmp_manualUpReq : BOOL;
    tmp_manualLeftReq : BOOL;
    tmp_manualRightReq : BOOL;
    tmp_manualGripReq : BOOL;
    tmp_manualReleaseReq : BOOL;

    tmp_autoDown : BOOL;
    tmp_autoUp : BOOL;
    tmp_autoLeft : BOOL;
    tmp_autoRight : BOOL;
    tmp_autoGrip : BOOL;
    tmp_autoRelease : BOOL;

    tmp_down : BOOL;
    tmp_up : BOOL;
    tmp_left : BOOL;
    tmp_right : BOOL;
    tmp_grip : BOOL;
    tmp_release : BOOL;
END_VAR

tmp_startEdge(CLK := Start);

tmp_manualDownReq := ManualMode AND DownButton AND NOT DownLimitSwitch;
tmp_manualUpReq := ManualMode AND UpButton AND NOT UpLimitSwitch;
tmp_manualLeftReq := ManualMode AND LeftButton AND NOT LeftLimitSwitch;
tmp_manualRightReq := ManualMode AND RightButton AND NOT RightLimitSwitch;
tmp_manualGripReq := ManualMode AND GripButton AND NOT GripLimitSwitch;
tmp_manualReleaseReq := ManualMode AND ReleaseButton AND NOT ReleaseLimitSwitch;

tmp_autoMode := SingleStepMode OR SingleCycleMode OR ContinuousMode;

IF EmergencyStop AND tmp_startEdge.Q THEN
    IF SingleStepMode THEN
        IF NOT tmp_autoActive THEN
            tmp_currentStep := tmp_singleNextStep;
            tmp_singleNextStep := (tmp_singleNextStep + 1) MOD 8;
            tmp_autoActive := TRUE;
        END_IF;
    ELSIF SingleCycleMode THEN
        IF NOT tmp_autoActive THEN
            tmp_currentStep := 0;
            tmp_autoActive := TRUE;
        END_IF;
    ELSIF ContinuousMode THEN
        IF NOT tmp_autoActive THEN
            tmp_currentStep := 0;
            tmp_autoActive := TRUE;
        END_IF;
    END_IF;
END_IF;

CASE tmp_currentStep OF
    0, 4:
        tmp_targetReached := DownLimitSwitch;
    1:
        tmp_targetReached := GripLimitSwitch;
    2, 6:
        tmp_targetReached := UpLimitSwitch;
    3:
        tmp_targetReached := RightLimitSwitch;
    5:
        tmp_targetReached := ReleaseLimitSwitch;
    7:
        tmp_targetReached := LeftLimitSwitch;
ELSE
    tmp_targetReached := FALSE;
END_CASE;

tmp_autoDown := tmp_autoMode AND tmp_autoActive AND ((tmp_currentStep = 0) OR (tmp_currentStep = 4)) AND NOT DownLimitSwitch;
tmp_autoGrip := tmp_autoMode AND tmp_autoActive AND (tmp_currentStep = 1) AND NOT GripLimitSwitch;
tmp_autoUp := tmp_autoMode AND tmp_autoActive AND ((tmp_currentStep = 2) OR (tmp_currentStep = 6)) AND NOT UpLimitSwitch;
tmp_autoRight := tmp_autoMode AND tmp_autoActive AND (tmp_currentStep = 3) AND NOT RightLimitSwitch;
tmp_autoRelease := tmp_autoMode AND tmp_autoActive AND (tmp_currentStep = 5) AND NOT ReleaseLimitSwitch;
tmp_autoLeft := tmp_autoMode AND tmp_autoActive AND (tmp_currentStep = 7) AND NOT LeftLimitSwitch;

tmp_down := tmp_manualDownReq OR tmp_autoDown;
tmp_up := tmp_manualUpReq OR tmp_autoUp;
tmp_left := tmp_manualLeftReq OR tmp_autoLeft;
tmp_right := tmp_manualRightReq OR tmp_autoRight;
tmp_grip := tmp_manualGripReq OR tmp_autoGrip;
tmp_release := tmp_manualReleaseReq OR tmp_autoRelease;

MoveDown := tmp_down AND NOT tmp_up AND EmergencyStop;
MoveUp := tmp_up AND NOT tmp_down AND EmergencyStop;
MoveLeft := tmp_left AND NOT tmp_right AND EmergencyStop;
MoveRight := tmp_right AND NOT tmp_left AND EmergencyStop;
ActivateGrip := tmp_grip AND NOT tmp_release AND EmergencyStop;
ActivateRelease := tmp_release AND NOT tmp_grip AND EmergencyStop;

IF EmergencyStop AND tmp_autoMode AND tmp_autoActive AND tmp_targetReached THEN
    IF SingleStepMode THEN
        tmp_autoActive := FALSE;
    ELSIF SingleCycleMode THEN
        IF tmp_currentStep >= 7 THEN
            tmp_autoActive := FALSE;
            tmp_currentStep := 0;
        ELSE
            tmp_currentStep := tmp_currentStep + 1;
        END_IF;
    ELSIF ContinuousMode THEN
        IF tmp_currentStep >= 7 THEN
            tmp_currentStep := 0;
        ELSE
            tmp_currentStep := tmp_currentStep + 1;
        END_IF;
    END_IF;
END_IF;

END_FUNCTION_BLOCK
